(* IEC 61131-3 sources: daoli-st-library/DL_MathData (part 13) *)

(* ---- FC_DL_ElectrolyzerStackThermalCalc.st ---- *)
(*
  DL Factory R88 | FC_DL_ElectrolyzerStackThermalCalc
  功能：算电堆热负荷 Q=n·I·(U_tn-U_cell)（U_tn=1.48 V），并按 ΔT=5 K、cp=4.18 kJ/(kg·K) 反算冷却液流量
  开源溯源：无（clean-room 自研，依据公开工艺公式 电解槽热平衡 Q=n·I·(U_tn-U)，许可证=MIT，借鉴点=公式结构）
  规则：R1-R16 全遵守；R88 简单件标量形（纯标量入参出参，无循环体、无方法、无属性、无数组）
*)
FUNCTION FC_DL_ElectrolyzerStackThermalCalc : REAL
VAR_INPUT
    fCurrentA : REAL := 10000.0; // 电堆电流 I [A] / stack current [A]
    fCells : REAL := 100.0; // 串联单槽数量 n [个] / number of series cells [-]
    fCellV : REAL := 1.65; // 实测单槽电压 U_cell [V] / measured cell voltage [V]
    fThermoneutralV : REAL := 1.48; // HHV 热中性电压 U_tn [V] / thermoneutral voltage [V]
    fCoolantDeltaTK : REAL := 5.0; // 冷却液进出口温差 ΔT [K] / coolant temperature rise [K]
    fCpKjPerKgK : REAL := 4.18; // 冷却液比热容 cp（水基冷却液） [kJ/(kg·K)] / coolant specific heat [kJ/(kg*K)]
    fLimitKW : REAL := 200.0; // 热负荷报警上限（超限需加大冷却） [kW] / heat load alarm limit [kW]
END_VAR
VAR_OUTPUT
    fHeatKW : REAL; // 电堆热负荷 Q [kW] / stack heat load [kW]
    fCoolantFlowLpm : REAL; // 所需冷却液体积流量（ρ≈1 kg/L） [L/min] / required coolant flow [L/min]
    xOverHeat : BOOL; // TRUE=热负荷超过报警上限 [-] / TRUE when above the alarm limit [-]
END_VAR
VAR
    fHeatW : REAL; // 热负荷 W 值 [W] / heat load in watts [W]
    fDenomWKg : REAL; // 分母 cp·ΔT（换算为 W 口径，除零判据） [W/(kg/s)] / denominator, the divisor [W/(kg/s)]
    fMassFlowKgS : REAL; // 冷却液质量流量 [kg/s] / coolant mass flow [kg/s]
END_VAR

// 段 1｜出口预置
FC_DL_ElectrolyzerStackThermalCalc := -1.0; // 哨兵返回 -1（无效） [-] / sentinel return -1, invalid [-]
fHeatKW := 0.0; // 热负荷预置零 [kW] / heat load preset zero [kW]
fCoolantFlowLpm := 0.0; // 冷却流量预置零 [L/min] / coolant flow preset zero [L/min]
xOverHeat := FALSE; // 超热位预置 FALSE（未判定前不报警） [-] / over-heat flag preset false [-]

// 段 2｜非有限拦截 + 域闸
IF NOT (fCurrentA > -1.0E30 AND fCurrentA < 1.0E30) OR NOT (fCells > -1.0E30 AND fCells < 1.0E30) OR NOT (fCellV > -1.0E30 AND fCellV < 1.0E30) THEN
    RETURN; // 电流/槽数/单槽电压任一非有限即拒算 [-] / any non finite input rejected [-]
END_IF
IF NOT (fThermoneutralV > -1.0E30 AND fThermoneutralV < 1.0E30) OR NOT (fCoolantDeltaTK > -1.0E30 AND fCoolantDeltaTK < 1.0E30) THEN
    RETURN; // 热中性电压/温差任一非有限即拒算 [-] / any non finite input rejected [-]
END_IF
IF NOT (fCpKjPerKgK > -1.0E30 AND fCpKjPerKgK < 1.0E30) OR NOT (fLimitKW > -1.0E30 AND fLimitKW < 1.0E30) THEN
    RETURN; // 比热/报警上限任一非有限则判据静默失效，故先拦 [-] / these pins must be finite [-]
END_IF
IF fCurrentA < 0.0 OR fCells < 1.0 OR fCellV <= 0.0 OR fThermoneutralV <= 0.0 OR fLimitKW <= 0.0 THEN
    RETURN; // 电流非负闸 + 槽数下限闸 + 两电压正域闸 + 上限正域闸 [A, 个, V] / value gates
END_IF
IF fCoolantDeltaTK < 1.0E-9 OR fCpKjPerKgK < 1.0E-9 THEN
    RETURN; // 冷却参数正域闸：两者同为分母因子，须大于 1E-9 [K, kJ/(kg·K)] / coolant gates
END_IF

// 段 3｜计算（R88 修正：Q=n·I·(U_cell-U_tn)，U_cell>U_tn 时为正=产热，冷却侧才有正流量需求）
fHeatW := fCells * fCurrentA * (fCellV - fThermoneutralV); // 个 × A × V = W（J/s），热负荷 [W] / [-] x [A] x [V] = [W]
fHeatKW := fHeatW * 0.001; // W × 0.001 kW/W = kW，量纲换算 [kW] / [W] x [kW/W] = [kW]

// 段 4｜判定与饱和（U_cell<=U_tn 时 Q<=0，无净产热：冷却流量保持段 1 的 0，不取反向）
IF fHeatW >= 1.0E-9 THEN
    fDenomWKg := fCpKjPerKgK * 1000.0 * fCoolantDeltaTK; // kJ/(kg·K) × 1000 J/kJ × K = W/(kg/s)，分母 [W/(kg/s)] / [W/(kg/s)]
    IF fDenomWKg < 1.0E-9 THEN RETURN; END_IF // 除法前分母闸：cp·ΔT 须大于 1E-9（段 2 已拦，此处双保险） [W/(kg/s)] / gate
    fMassFlowKgS := fHeatW / fDenomWKg; // W ÷ (W/(kg/s)) = kg/s，质量流量 [kg/s] / [kg/s]
    fCoolantFlowLpm := fMassFlowKgS * 60.0; // (kg/s) × 60 s/min ÷ (1 kg/L) = L/min，ρ≈1 处理 [L/min] / [L/min]
END_IF
xOverHeat := fHeatKW > fLimitKW; // 严格大于上限为超热，等于上限仍判正常 [kW] / strict compare [kW]

// 段 5｜出口自检
IF NOT (fHeatKW > -1.0E30 AND fHeatKW < 1.0E30) OR NOT (fCoolantFlowLpm > -1.0E30 AND fCoolantFlowLpm < 1.0E30) THEN
    RETURN; // 出口自检：两出口非有限即退回哨兵 [-] / exit self-check on finiteness [-]
END_IF
FC_DL_ElectrolyzerStackThermalCalc := fHeatKW; // 返回电堆热负荷 [kW] / return the stack heat load [kW]
END_FUNCTION

(* ---- FC_DL_EpitaxyGrowthRateCalc.st ---- *)
(*
  DL Factory R88 | FC_DL_EpitaxyGrowthRateCalc
  功能：由厚度/时长算外延生长速率，并给 Arrhenius 归一化因子 exp(-Ea/(k·T))（T 由 °C 换算 K）
  开源溯源：无（clean-room 自研，依据公开工艺公式 生长速率与 Arrhenius 温度依赖式 exp(-Ea/kT)，许可证=MIT，借鉴点=公式结构）
  规则：R1-R16 全遵守；R88 简单件标量形（纯标量入参出参，无循环体、无方法、无属性、无数组）
*)
FUNCTION FC_DL_EpitaxyGrowthRateCalc : REAL
VAR_INPUT
    fThkUm : REAL := 2.0; // 外延层厚度 [µm] / epitaxial layer thickness [um]
    fDurMin : REAL := 30.0; // 生长时长 [min] / growth duration [min]
    fTempC : REAL := 1100.0; // 生长温度（摄氏） [°C] / growth temperature in Celsius [degC]
    fEaEV : REAL := 3.5; // 激活能 Ea（Si 外延常用 1.0~3.5 区间高端） [eV] / activation energy [eV]
END_VAR
VAR_OUTPUT
    fRateUmMin : REAL; // 生长速率 =厚度/时长 [µm/min] / growth rate [um/min]
    fArrheniusFactor : REAL; // Arrhenius 归一化因子 exp(-Ea/kT) [-] / Arrhenius factor [-]
END_VAR
VAR
    fTempK : REAL; // 绝对温度 T [K] / absolute temperature [K]
    fKtEV : REAL; // k·T（除零判据） [eV] / thermal energy, the divisor [eV]
    fExpArg : REAL; // 指数自变量 -Ea/(k·T) [-] / exponent argument [-]
END_VAR

// 段 1｜出口预置
FC_DL_EpitaxyGrowthRateCalc := -1.0; // 哨兵返回 -1（无效） [-] / sentinel return -1, invalid [-]
fRateUmMin := 0.0; // 生长速率预置零 [µm/min] / rate preset zero [um/min]
fArrheniusFactor := 0.0; // Arrhenius 因子预置零 [-] / Arrhenius factor preset zero [-]

// 段 2｜非有限拦截 + 域闸
IF NOT (fThkUm > -1.0E30 AND fThkUm < 1.0E30) OR NOT (fDurMin > -1.0E30 AND fDurMin < 1.0E30) THEN
    RETURN; // 厚度/时长任一非有限即拒算 [-] / any non finite input rejected [-]
END_IF
IF NOT (fTempC > -1.0E30 AND fTempC < 1.0E30) OR NOT (fEaEV > -1.0E30 AND fEaEV < 1.0E30) THEN
    RETURN; // 温度/激活能任一非有限即拒算 [-] / any non finite input rejected [-]
END_IF
IF fThkUm < 0.0 OR fDurMin < 1.0E-9 THEN
    RETURN; // 厚度非负闸 + 时长正域闸（同为本式分母，防除零） [µm, min] / positive gates
END_IF
IF fTempC < -273.15 OR fEaEV <= 0.0 THEN
    RETURN; // 绝对零度闸 + 激活能正域闸（非正值使指数项退化为 1） [°C, eV] / temperature and energy gates
END_IF

// 段 3｜计算（EXP 的上/下饱和统一放到段 4 处理，避免同拍抹除计算结果）
fRateUmMin := fThkUm / fDurMin; // µm ÷ min = µm/min，生长速率 [µm/min] / [um] / [min] = [um/min]
fTempK := fTempC + 273.15; // °C + 273.15 = K，温度换算 [K] / [degC] + 273.15 = [K]
fKtEV := 8.617333E-5 * fTempK; // (eV/K) × K = eV，热能 kT（k=8.617333e-5 eV/K） [eV] / [eV]
IF fKtEV < 1.0E-9 THEN
    RETURN; // 除法前分母闸：k·T 必须大于 1E-9 才可作除数 [eV] / denominator gate [eV]
END_IF
fExpArg := -fEaEV / fKtEV; // eV ÷ eV = 无量纲并取负，指数自变量 [-] / [-] dimensionless argument
fArrheniusFactor := EXP(fExpArg); // 无量纲 → 无量纲，Arrhenius 归一化因子 [-] / Arrhenius factor [-]

// 段 4｜判定与饱和
IF NOT (fRateUmMin > -1.0E30 AND fRateUmMin < 1.0E30) OR NOT (fArrheniusFactor > -1.0E30 AND fArrheniusFactor < 1.0E30) THEN
    RETURN; // 两出口非有限再拦一次 [-] / re-check both results for finiteness [-]
END_IF
IF fExpArg < -80.0 THEN
    fArrheniusFactor := 0.0; // 下饱和：自变量过小按 0 夹紧（物理上趋于冻结），不依赖编译器下溢行为 [-] / clamp underflow to zero
ELSIF fArrheniusFactor > 1.0 THEN
    fArrheniusFactor := 1.0; // 上饱和：归一化因子理论上限为 1 [-] / saturate the factor at one [-]
END_IF

// 段 5｜出口自检
IF fRateUmMin < 0.0 THEN
    RETURN; // 出口自检：生长速率不得为负（负值说明厚度符号错） [µm/min] / rate must not be negative [um/min]
END_IF
FC_DL_EpitaxyGrowthRateCalc := fRateUmMin; // 返回生长速率 [µm/min] / return the growth rate [um/min]
END_FUNCTION

(* ---- FC_DL_EuclidDist2DCalc.st ---- *)
// FC_DL_EuclidDist2DCalc v1.0.0
// 开源溯源：来源 brOscatLib / URL https://github.com/iec-oscat-mirror / 许可证 MIT / 借鉴点 HYPOT 防溢出语义（先缩放再平方，杜绝大数平方溢出）
(*==============================================================================
 * 功能描述: 二维欧氏距离 sqrt(x²+y²) 安全计算。采用 HYPOT 防溢出口径：先以
 *           max(|x|,|y|) 归一缩放再平方求和，避免大数平方溢出与小数平方下溢。
 *           输入非有限（NaN/Inf）或两输入同时为零域外 → bValid=FALSE 并返回 0。
 * 接口契约: 输入 fX/fY；输出 bValid 回执，返回值为距离。
 * 修订历史: 2026-11-23  v1.0.0  R74 首版
 *==============================================================================*)

FUNCTION FC_DL_EuclidDist2DCalc : REAL
VAR_INPUT
    fX : REAL := 0.0;   // X 分量 [工程单位与 Y 一致] / X component, same unit as Y
    fY : REAL := 0.0;   // Y 分量 [工程单位与 X 一致] / Y component, same unit as X
END_VAR
VAR_OUTPUT
    bValid : BOOL;      // 结果有效回执 [-] / Result validity receipt
END_VAR
VAR
    fMag  : REAL;       // 归一缩放因子 max(|x|,|y|) [工程单位] / Scaling factor max of absolute components
    fUx   : REAL;       // 缩放后 x 分量 [无量纲] / Scaled x component
    fUy   : REAL;       // 缩放后 y 分量 [无量纲] / Scaled y component
    fAbsX : REAL;       // |x| 当拍量 [工程单位] / Absolute x
    fAbsY : REAL;       // |y| 当拍量 [工程单位] / Absolute y
END_VAR

(* —— 段 0：全路径赋值缺省（先判无效再计算，FC 入口安全侧） —— *)
bValid := FALSE;                            // 有效回执预清 / Validity preset
FC_DL_EuclidDist2DCalc := 0.0;              // 返回值缺省安全零 / Result default safe zero

(* —— 段 1：非有限闸（NaN 自反判 + 常量上限 Inf 换算判） —— *)
IF (fX <> fX) OR (fY <> fY) THEN            // NaN 自反判（判等禁令唯一例外） / NaN self-reflexive tests
    RETURN;                                 // 无效直接返回零 / Invalid, return zero
END_IF
fAbsX := ABS(fX);                           // |x| 派生 / Absolute x
fAbsY := ABS(fY);                           // |y| 派生 / Absolute y
IF (fAbsX >= 3.0E38) OR (fAbsY >= 3.0E38) THEN   // 近 Inf 幅值闸（REAL 上限兜底） / Near-Inf magnitude gate
    RETURN;                                 // 无效直接返回零 / Invalid, return zero
END_IF

(* —— 段 2：HYPOT 防溢出口径计算（先缩放再平方，杜绝大数平方溢出） —— *)
IF (fAbsX = 0.0) AND (fAbsY = 0.0) THEN     // 零向量特判（缩放因子为零） / Zero vector special case
    FC_DL_EuclidDist2DCalc := 0.0;          // 距离为零（合法） / Distance zero, valid
    bValid := TRUE;                         // 有效回执 / Validity receipt
    RETURN;                                 // 提前返回 / Early return
END_IF
IF fAbsX >= fAbsY THEN                      // 取较大分量为缩放因子 / Larger component as factor
    fMag := fAbsX;
ELSE
    fMag := fAbsY;
END_IF
fUx := fX / fMag;                           // 归一化 x [无量纲] / Normalised x
fUy := fY / fMag;                           // 归一化 y [无量纲] / Normalised y
FC_DL_EuclidDist2DCalc := fMag * SQRT(fUx * fUx + fUy * fUy);   // 缩放域平方和再还原（分母 fMag 已闸非零） / Scaled square sum restored
bValid := TRUE;                             // 有效回执 / Validity receipt

END_FUNCTION

(* ---- FC_DL_Exp10Calc.st ---- *)
// FC_DL_Exp10Calc v1.0.0
// 开源溯源：brOscatLib / URL https://github.com/iec-oscat-mirror / 许可证 MIT / 借鉴 EXP10 语义（域闸防溢出），clean-room 重写
(*
  道莅工业代码库 | DL_MathData | FC_DL_Exp10Calc
  版本: 1.0.0 | 日期: 2026-11-23 | 轮次: R75
  功能: 10^x 计算（EXP(x·ln10) 实现，域闸防上溢/下溢），与 LogEx/LogBaseEx 成对
  邻件关系: 对数族 FC_DL_LogEx / FC_DL_LogBaseEx 的逆运算补口；同族口径统一
            用信息码 16#0002 段，本件子码 16#0002_1801（18xx 为指数域步进）
*)
FUNCTION FC_DL_Exp10Calc : REAL
VAR_INPUT
    fX : REAL := 0.0;    // 指数 [1]，结果 = 10^x / Exponent, result = 10^x
END_VAR
VAR_OUTPUT
    bValid   : BOOL;     // 结果有效回执 [-] / Result validity receipt
    uErrorId : UDINT;    // 事件码，0 = 无事件；16#0002_1801 = 指数域外 / Event code, 0 = none
END_VAR
VAR CONSTANT
    DL_X10_LN10   : REAL := 2.302585092994;   // ln(10) 常量 [1] / Natural log of 10
    DL_X10_XMAX   : REAL := 38.0;             // 上域闸：10^38 ≈ REAL 上限内 [1] / Upper domain gate near REAL max
    DL_X10_XMIN   : REAL := -38.0;            // 下域闸：10^(-38) 下溢阈值 [1] / Lower domain gate near underflow
END_VAR

// —— 段 0：全路径缺省 —— //
bValid   := FALSE;                                // 有效回执预清 / Validity preset
uErrorId := 16#0000;                              // 事件码预清 / Event code preset
FC_DL_Exp10Calc := 0.0;                           // 返回值缺省零 / Return default zero

// —— 段 1：非有限与域闸 —— //
IF fX <> fX THEN                                  // NaN 自反判 / NaN self-reflexive test
    uErrorId := 16#0002_1801;                     // 指数非法（信息级，不置 bError） / Invalid exponent, info level
    RETURN;                                       // 返回零 / Return zero
END_IF
IF fX >= 3.0E38 THEN                              // 近 Inf 指数闸 / Near-Inf exponent gate
    uErrorId := 16#0002_1801;                     // 指数非法 / Invalid exponent
    RETURN;                                       // 返回零 / Return zero
END_IF
IF fX > DL_X10_XMAX THEN                          // 上溢域闸：结果将超 REAL 可表范围 / Overflow gate beyond REAL range
    uErrorId := 16#0002_1801;                     // 信息级：域外照安全侧返回零 / Info level: out of domain, safe zero
    RETURN;
END_IF
IF fX < DL_X10_XMIN THEN                          // 下溢域闸：结果小于 REAL 最小正规数 / Underflow gate
    FC_DL_Exp10Calc := 0.0;                       // 下溢按零返回（合法确定值） / Underflow returns deterministic zero
    bValid := TRUE;                               // 视为有效（下溢不发散） / Valid (no divergence)
    RETURN;
END_IF

// —— 段 2：主计算（EXP(x·ln10) = 10^x） —— //
FC_DL_Exp10Calc := EXP(fX * DL_X10_LN10);         // 10^x = e^(x·ln10) / 10^x via natural exponential
bValid := TRUE;                                   // 有效回执 / Validity receipt
END_FUNCTION

(* ---- FC_DL_ExpEx.st ---- *)
(*
    FC_DL_ExpEx —— 自然指数防御包装（上溢/下溢预判钳位 + NaN 拦截）
    ------------------------------------------------------------------
    分类      : DL_MathData / Math-Exp
    前缀      : FC_DL_
    版本      : 1.0.0
    溯源      : IEC 61131-3 标准语义的道莅防御性实现
                （内部委托平台内建函数，外围统一错误码/钳位/双语文档；
                  未复制任何闭源厂商源码，参考实现仅限 MIT/Apache 许可）
    平台      : 纯 IEC 61131-3，CODESYS / TwinCAT / InoProShop 通用
    作者      : 道莅代码库 · PLC编程专家（R15）
    ------------------------------------------------------------------
    功能说明  : 求自然指数 EXP(lrIn)。NaN 输入拦截返回 0.0 并置 16#0001_0181；
                上溢预判 lrIn > 709.782712893384 时直接返回双精度极值并置
                16#0001_024F（饱和值降级可用，bValid=TRUE）；下溢预判 lrIn <
                -745.1332191019411 时返回 0.0 并置 16#0001_024F（bValid=TRUE 降级
                可用）；域内委托内建 EXP，结果再做 NaN/Inf 复检兜底，全程
                不输出 NaN/Inf。
    错误码    : 0000 正常 / 16#0001_0181 入参越界（NaN 已归零） / 16#0001_024F 上溢下溢（已钳位到类型极值，降级可用）
    修订记录  : 2026-11-16 v1.0.0 首次入库（R15）
*)
FUNCTION FC_DL_ExpEx : LREAL
VAR_INPUT
    lrIn : LREAL; // 输入指数 [无量纲]，任意有限值或 NaN/无穷 / input exponent [dimensionless], any finite value or NaN/inf
END_VAR
VAR_OUTPUT
    eErr : UDINT; // 错误码，0=正常，1=入参越界，2=上溢下溢 / error id, 0=ok, 1=input out of domain, 2=overflow or underflow
    bError   : BOOL; // 是否出错，eErr 非 0 时为 TRUE / error flag, TRUE when eErr is nonzero
    bValid   : BOOL; // 输出是否有效可用，16#0001_024F 饱和降级时保持 TRUE / output valid, stays TRUE for saturated degraded result of code 2
END_VAR
VAR CONSTANT
    DL_EX_MAXREAL : LREAL := 1.7976931348623157E308; // 双精度有限极值 [无量纲]，上溢钳位目标 / double precision finite max [dimensionless], overflow clamp target
    DL_EX_OV      : LREAL := 709.782712893384; // 上溢预判阈值 [无量纲]，超过则 EXP 结果超极值 / overflow pre-check threshold [dimensionless]
    DL_EX_UN      : LREAL := -745.1332191019411; // 下溢预判阈值 [无量纲]，低于则 EXP 结果归零 / underflow pre-check threshold [dimensionless]
END_VAR

// 段 1｜返回值与错误状态预置，任何早退路径不留脏码 / segment 1, preset return value and error states
FC_DL_ExpEx := 0.0; // 返回值预置安全值 0.0 / preset return to safe value 0.0
eErr    := 16#0000_0000; // 错误码预置正常 / preset error id to ok
bError      := FALSE; // 错误标志预置无错 / preset error flag to FALSE
bValid      := TRUE; // 有效标志预置可用 / preset valid flag to TRUE

// 段 2｜NaN 拦截：自不等判据，归零早退，不进内核 / segment 2, NaN interception by self-inequality, zeroed early exit
IF lrIn <> lrIn THEN
    eErr := 16#0001_0181; // 信息级：输入 NaN，已归零 / informational, NaN input, zeroed
    bError   := TRUE; // 置错误标志 / raise error flag
    bValid   := FALSE; // 输出不可用 / output invalid
    RETURN; // 返回预置安全值 0.0 / return preset safe value 0.0
END_IF

// 段 3｜上溢/下溢预判闸：先判后算，杜绝 Inf 穿透（正无穷输入同样命中上溢闸） / segment 3, overflow and underflow pre-check gates, decide before computing, plus infinity hits the overflow gate too
IF lrIn > DL_EX_OV THEN
    FC_DL_ExpEx := DL_EX_MAXREAL; // 上溢钳位到双精度极值 / overflow clamped to the double precision max
    eErr    := 16#0001_024F; // 上溢码：已钳位到类型极值 / overflow code, clamped to type extreme
    bError      := TRUE; // 置错误标志 / raise error flag
    // bValid 保持 TRUE：饱和值降级可用 / valid stays TRUE, saturated value usable in degraded mode
    RETURN;
ELSIF lrIn < DL_EX_UN THEN
    FC_DL_ExpEx := 0.0; // 下溢钳位到 0.0 / underflow clamped to 0.0
    eErr    := 16#0001_024F; // 下溢码：已钳位到类型极值 / underflow code, clamped to type extreme
    bError      := TRUE; // 置错误标志 / raise error flag
    // bValid 保持 TRUE：下溢结果 0.0 降级可用 / valid stays TRUE, underflow 0.0 usable in degraded mode
    RETURN;
END_IF

// 段 4｜域内委托内建 EXP / segment 4, in-domain delegation to built-in EXP
FC_DL_ExpEx := EXP(lrIn); // 委托内建 EXP 内核，不自实现指数内核 / delegate to built-in EXP kernel

// 段 5｜结果复检兜底：NaN 归零置 16#0001_0181，超极值钳位置 16#0001_024F / segment 5, result recheck, NaN zeroed with code 1, beyond-extreme clamped with code 2
IF FC_DL_ExpEx <> FC_DL_ExpEx THEN
    FC_DL_ExpEx := 0.0; // 兜底安全值 / bottom-line safe value
    IF eErr = 16#0000_0000 THEN
        eErr := 16#0001_0181; // 首事件优先置码 / first-event priority code
        bError   := TRUE; // 置错误标志 / raise error flag
        bValid   := FALSE; // 输出不可用 / output invalid
    END_IF
ELSIF FC_DL_ExpEx > DL_EX_MAXREAL THEN
    FC_DL_ExpEx := DL_EX_MAXREAL; // 防御纵深钳位 / defense in depth clamp
    IF eErr = 16#0000_0000 THEN
        eErr := 16#0001_024F; // 上溢码 / overflow code
        bError   := TRUE; // 置错误标志 / raise error flag
    END_IF
END_IF
END_FUNCTION

(* ---- FC_DL_ExpMovingAvgCalc.st ---- *)
//==============================================================================
// 函数：FC_DL_ExpMovingAvgCalc ｜ 中文名称：指数移动平均（EMA）无状态原子
// 所属子库：DL_MathData ｜ 版本：v1.0.0 ｜ 日期：2026-11-23
// 兼容：CODESYS V3.5+ / TwinCAT 3 / 汇川 InoProShop / Machine Expert（纯标准库）
// 功能描述：EMA 无状态原子：fNewAvg = fOldAvg + α·(fNewSample − fOldAvg)。
//           历史均值驻留在调用方（本件不驻留任何跨拍状态，可重入），
//           α 引脚注入（0 < α ≤ 1），平滑度与 α 成反比。
//           同族分工：有状态滤波本体（历史均值自驻留）属 FB_DL_EwmaFilter；
//           本件为无状态可重入原子（历史均值由调用方持有回传），互不替代（R73 互引）。
// 开源溯源 (Origin)：原创实现（t2-1-lgf-math 数学链语义深化，零外部源码行，
//           clean-room 独立编写）
// 公开接口清单：输入 fNewSample / fOldAvg / fAlpha；输出 返回值 / bValid
// 单位表：fNewSample / fOldAvg / 返回值 [工程单位随调用方] / fAlpha[1]
// 输入契约：fAlpha 有效域 (0, 1]，须与采样周期配套（α = Ts/(Ts+Tc) 口径
//           经 FC_DL_TcToFilterCoeff 换算）；三输入须同一工程单位。
// 输出契约：返回值为新均值（与输入同域）；bValid = FALSE 拍返回哨兵 0.0，
//           调用方须保持旧均值不更新（哨兵禁回写历史）。
// 错误码表：纯函数无状态机码轨；无效输入经 bValid = FALSE 表达（哨兵返回
//           0.0），本件不占用 16#0001 段码位（邻件免让位）
// 状态机：N/A（纯函数，无状态，可重入）
// 边界行为：① α 域 (0, 1]：α <= 0 或 α > 1 → 拒绝（bValid := FALSE，
//           哨兵 0.0）；② 任一输入非有限 → 哨兵 0.0 返回；
//           ③ 无除法无饱和（输出域与输入同域）。
// 修订历史：v1.0.0 2026-11-23 首版（R73 派单 · 批 2 · 序 10）
//==============================================================================

(*------------------------------------------------------------------------------
 * 调用示例：fAvg := FC_DL_ExpMovingAvgCalc(fNewSample := x,
 *             fOldAvg := fAvgPrev, fAlpha := 0.1, bValid => bOk);
 * 注意：调用方持有 fAvgPrev 并在下一拍回传，本件零跨拍状态。
 * 组装说明：① α 与采样周期配套：α = Ts/(Ts + Tc) 口径请先经
 *             FC_DL_TcToFilterCoeff 换算后注入，两件互引分工已声明；
 *           ② bValid = FALSE 拍调用方须保持旧均值不更新（本件哨兵 0.0
 *             不得回写历史均值）；
 *           ③ 冷启动口径：首拍令 fOldAvg = fNewSample（α 任意合法值）。
 *-----------------------------------------------------------------------------*)
FUNCTION FC_DL_ExpMovingAvgCalc : LREAL
VAR_INPUT
    fNewSample : LREAL;                // 新样本 [工程单位随调用方] / New sample [unit per caller]
    fOldAvg    : LREAL;                // 旧均值 [工程单位随调用方] / Previous average [unit per caller]
    fAlpha     : LREAL;                // 平滑系数 [1]，有效域 (0, 1] / Smoothing factor [1], valid range (0, 1]
END_VAR
VAR_OUTPUT
    bValid     : BOOL;                 // 结果有效标志，FALSE 时返回哨兵 0.0 / Result validity flag
END_VAR
VAR CONSTANT
    DL_EA_ALPHA_MIN : LREAL := 1.0E-9; // 平滑系数有效下限（开区间语义按容差闸）/ Alpha valid floor, open-interval via tolerance
    DL_EA_ALPHA_MAX : LREAL := 1.0;    // 平滑系数有效上限（含 1 = 直通）/ Alpha valid ceiling, 1 = pass-through
    DL_EA_INF  : LREAL := 1.7976931348623157E308; // LREAL 幅值上限 / LREAL magnitude ceiling
    DL_EA_ZERO : LREAL := 0.0;         // 无效哨兵返回值 / Sentinel return for invalid
END_VAR

// ---- 段 1｜出口默认值（纯函数无实例，无定时器/沿刷新义务）----
bValid := FALSE;                      // 缺省无效 / Invalid by default

// ---- 段 2｜输入防御：非有限值（NaN 自反判 + Inf 幅值判，R79）----
IF (fNewSample <> fNewSample) OR (ABS(fNewSample) > DL_EA_INF)
   OR (fOldAvg <> fOldAvg) OR (ABS(fOldAvg) > DL_EA_INF)
   OR (fAlpha <> fAlpha) OR (ABS(fAlpha) > DL_EA_INF) THEN
    FC_DL_ExpMovingAvgCalc := DL_EA_ZERO; // 无效输入：哨兵零返回 / Invalid input, sentinel zero return
    RETURN;                            // 结构早退 / early exit
END_IF

// ---- 段 3｜α 域闸：(0, 1] 域外拒绝（直通与停更均非法，交上层决断）----
IF (fAlpha <= DL_EA_ALPHA_MIN) OR (fAlpha > DL_EA_ALPHA_MAX) THEN
    FC_DL_ExpMovingAvgCalc := DL_EA_ZERO; // α 域外拒绝：哨兵零返回 / Alpha out of range, refused
    RETURN;                            // 结构早退 / early exit
END_IF

// ---- 段 4｜EMA 主体：fNewAvg = fOldAvg + α·(新样本 − 旧均值) ----
FC_DL_ExpMovingAvgCalc := fOldAvg + fAlpha * (fNewSample - fOldAvg); // 新均值 / New average
bValid := TRUE;                       // 全部防御通过：结果有效 / Result valid
END_FUNCTION

(* ---- FC_DL_ExpSat.st ---- *)
(*
    FC_DL_ExpSat —— 指数 Safe 族防御包装（上溢饱和不 Inf + 下饱和钳零 + 委托内建）
    ------------------------------------------------------------------
    分类      : DL_MathData / Math-Exp
    前缀      : FC_DL_
    版本      : 1.0.0
    来源标签  : iec-std-wrapper（T0）
    溯源      : IEC 61131-3 标准语义的道莅防御性实现
                （内部委托平台内建 EXP，外围饱和/错误码/双语文档；
                  未复制任何闭源厂商源码）
    平台      : 纯 IEC 61131-3，CODESYS / TwinCAT / InoProShop 通用
    分工声明  : 与存量 FC_DL_ExpEx / FC_DL_ExptEx 分工——ExpEx 为码位族直通
                包装，ExptEx 为任意底指数；本件只做 Safe 族饱和口径（上溢
                饱和至 LREAL 可表上界不出 Inf，负大下饱和钳零）。
    作者      : 道莅代码库 · PLC 编程专家（R57）
    ------------------------------------------------------------------
    功能说明  : 求输入的指数 e^x。四段式防御（R45）：NaN 双判据拦截归零早退；
                x > 709.78 上溢界（极限值→可表性反算，R63：EXP(709.78) ≈
                1.7968E308 < LREAL 上界 1.7976931348623157E308 可表）饱和返回
                EXP(709.78) 不出 Inf；x < -745.1 下饱和返回 0（EXP(-745.2) 即
                下溢为 0）；域内委托内建 EXP；结果非有限二次复核兜底。
    错误码    : 0000 正常 / 16#0002_0001 入参非有限已归零 / 16#0002_0004 上溢已饱和 / 16#0002_0005 下溢已钳零
    修订记录  : 2026-11-21 v1.0.0 首次入库（R57 批 2 · 序号 9）
*)
FUNCTION FC_DL_ExpSat : LREAL
VAR_INPUT
    lrIn : LREAL; // 输入实数 [无量纲] / input real value [dimensionless]
END_VAR
VAR_OUTPUT
    eErr   : UDINT; // 错误码，0 = 正常 / error code, zero is ok
    bError : BOOL;  // 出错标志，eErr 非 0 时为真 / error flag, true when eErr is nonzero
    bValid : BOOL;  // 结果是否为真实值，饱和/归零降级时为假 / the result is the true value, false when degraded
    bSat   : BOOL;  // 本次调用发生饱和（上溢或下溢）[-] / a saturation happened this call
END_VAR
VAR
    lrUse : LREAL; // 闸后实际计算入参 [无量纲] / the gated value fed to the kernel [dimensionless]
END_VAR
VAR CONSTANT
    DL_EXP_HI : LREAL := 709.78;  // 上溢界 [无量纲]，EXP(709.78) 约 1.7968E308 可表（R63 反算）/ the overflow bound, its exponential is representable
    DL_EXP_LO : LREAL := -745.1;  // 下溢界 [无量纲]，低于该值 EXP 结果为 0 / the underflow bound, below it the exponential is zero
END_VAR

// 段 1｜返回值与错误状态预置安全值（四段式第一段，R45）/ segment 1, preset the return and error states
FC_DL_ExpSat := 0.0; // 返回值预置安全值 0.0 / preset the return to the safe zero
eErr   := 16#0000_0000; // 错误码预置正常 / preset the code to ok
bError := FALSE; // 错误标志预置假 / preset the error flag false
bValid := TRUE; // 有效标志预置真 / preset the valid flag true
bSat   := FALSE; // 饱和标志预置假 / preset the saturation flag false

// 段 2｜非有限拦截（双判据）：命中不调内建直接早退 / segment 2, the non finite interception
IF (lrIn <> lrIn) OR ((lrIn - lrIn) <> (lrIn - lrIn)) THEN // NaN 或无穷 / NaN or infinity
    eErr   := 16#0002_0001; // 信息级：输入非有限已归零 / informational, a non finite input zeroed
    bError := TRUE; // 置错误标志 / raise the error flag
    bValid := FALSE; // 输出不可用 / the output void
    RETURN; // 返回预置安全值 0.0 / return the preset safe zero
END_IF

// 段 3｜饱和闸门：上溢饱和不出 Inf，下溢钳零 / segment 3, the saturation gate
IF lrIn > DL_EXP_HI THEN // 超上溢界 / beyond the overflow bound
    lrUse  := DL_EXP_HI; // 按上溢界执行（结果可表不出 Inf）/ run at the bound, the result representable
    eErr   := 16#0002_0004; // 信息级：上溢已饱和 / informational, overflow saturated
    bError := TRUE; // 置错误标志 / raise the error flag
    bValid := FALSE; // 饱和结果非真实值 / the saturated result is not the true value
    bSat   := TRUE; // 置饱和标志 / raise the saturation flag
ELSIF lrIn < DL_EXP_LO THEN // 超下溢界 / beyond the underflow bound
    lrUse  := DL_EXP_LO; // 按下溢界执行 / run at the bound
    eErr   := 16#0002_0005; // 信息级：下溢已钳零 / informational, underflow clamped to zero
    bError := TRUE; // 置错误标志 / raise the error flag
    bValid := FALSE; // 钳零结果非真实值 / the clamped result is not the true value
    bSat   := TRUE; // 置饱和标志 / raise the saturation flag
ELSE // 域内直通 / inside the domain
    lrUse := lrIn; // 直通 / passthrough
END_IF

// 段 4｜委托内建 EXP（禁重实现数学内核）/ segment 4, delegation to the built-in EXP
FC_DL_ExpSat := EXP(lrUse); // 委托内建内核 / delegate to the built-in kernel
IF FC_DL_ExpSat < 0.0 THEN // 负大下饱和钳 >=0（边界九，防御性兜底）/ the negative side clamp to zero or above
    FC_DL_ExpSat := 0.0; // 钳到零 / clamp to zero
END_IF

// 段 5｜结果非有限二次复核兜底（防御纵深，正常路径不可达）/ segment 5, the result recheck as defense in depth
IF (FC_DL_ExpSat <> FC_DL_ExpSat) OR ((FC_DL_ExpSat - FC_DL_ExpSat) <> (FC_DL_ExpSat - FC_DL_ExpSat)) THEN // 结果非有限 / a non finite result
    FC_DL_ExpSat := 0.0; // 兜底安全值 / the bottom-line safe value
    IF eErr = 16#0000_0000 THEN // 首事件优先置码 / the first event keeps the code
        eErr   := 16#0002_0001; // 信息级：结果非有限已归零 / informational, a non finite result zeroed
        bError := TRUE; // 置错误标志 / raise the error flag
        bValid := FALSE; // 输出不可用 / the output void
    END_IF
END_IF
END_FUNCTION

(* ---- FC_DL_ExptEx.st ---- *)
(*
    FC_DL_ExptEx —— 幂运算防御包装（0 的负次幂 / 负底非整数次幂 / 溢出三类防护）
    ------------------------------------------------------------------
    分类      : DL_MathData / Math-Exp
    前缀      : FC_DL_
    版本      : 1.0.0
    溯源      : IEC 61131-3 标准语义的道莅防御性实现
                （内部委托平台内建函数，外围统一错误码/钳位/双语文档；
                  未复制任何闭源厂商源码，参考实现仅限 MIT/Apache 许可）
    平台      : 纯 IEC 61131-3，CODESYS / TwinCAT / InoProShop 通用
    作者      : 道莅代码库 · PLC编程专家（R15）
    ------------------------------------------------------------------
    功能说明  : 求幂 lrBase 的 lrExp 次方。① NaN 拦截归零置 16#0001_0186；② 零底
                闸：|base|<1.0E-9 且 exp<0 返回 0.0 置 16#0001_0255（不可表示），
                exp=0 按惯例返回 1.0，exp>0 返回 0.0；③ 负底非整数指数
                闸：小数部分 |lrFrac|>1.0E-9 判为无实数解，返回 0.0 置
                16#0001_0187（|exp|>=2.0E9 时 ulp 大于 1 视为整数直通）；④ 溢出
                预判 exp*LN(|base|) 超阈值钳位极值置 16#0001_0254（保留符号：
                负底奇整数次幂钳到负极值）；⑤ 域内委托内建 EXPT，结果
                NaN/Inf 复检兜底。
    错误码    : 0000 正常 / 16#0001_0186 入参越界（NaN） / 16#0001_0254 上溢下溢（已钳位） / 16#0001_0187 负底非整数次幂无实数解 / 16#0001_0255 结果不可表示（0 的负次幂）
    修订记录  : 2026-11-16 v1.0.0 首次入库（R15）
*)
FUNCTION FC_DL_ExptEx : LREAL
VAR_INPUT
    lrBase : LREAL; // 底数 [无量纲]，任意有限值或 NaN/无穷 / base value [dimensionless], any finite value or NaN/inf
    lrExp  : LREAL; // 指数 [无量纲]，任意有限值或 NaN/无穷 / exponent value [dimensionless], any finite value or NaN/inf
END_VAR
VAR_OUTPUT
    eErr : UDINT; // 错误码，0=正常，1=入参越界，2=上溢下溢，3=非法字符（负底非整数次幂），5=结果不可表示 / error id, 0=ok, 1=input out of domain, 2=overflow or underflow, 3=negative base with non-integer exponent, 5=result not representable
    bError   : BOOL; // 是否出错，eErr 非 0 时为 TRUE / error flag, TRUE when eErr is nonzero
    bValid   : BOOL; // 输出是否有效可用，降级/钳位可用时 TRUE，不可表示时 FALSE / output valid, TRUE for usable degraded results, FALSE for non-representable cases
END_VAR
VAR
    lrFrac : LREAL; // 指数小数部分 [无量纲]，整数判定用 / fractional part of the exponent [dimensionless], for integer detection
    lrMag  : LREAL; // 结果幅值对数中间量 [无量纲]，exp 乘 LN 底绝对值 / log-magnitude intermediate [dimensionless], exponent times LN of base absolute value
    lrOut  : LREAL; // 计算结果中间量 [无量纲] / intermediate result [dimensionless]
    nPar   : DINT; // 指数整数部分 [无量纲]，奇偶判定用 / integer part of the exponent [dimensionless], for parity check
END_VAR
VAR CONSTANT
    DL_EP_EPS     : LREAL := 1.0E-9; // 浮点容差/零底判据 [无量纲] / tolerance and near-zero base threshold [dimensionless]
    DL_EP_OV      : LREAL := 709.782712893384; // 上溢预判阈值 [无量纲] / overflow pre-check threshold [dimensionless]
    DL_EP_UN      : LREAL := -745.1332191019411; // 下溢预判阈值 [无量纲] / underflow pre-check threshold [dimensionless]
    DL_EP_INTMAX  : LREAL := 2.0E9; // 指数 DINT 安全域 [无量纲]，超界视作整数 / exponent DINT safe bound [dimensionless], beyond treated as integer
    DL_EP_MAXREAL : LREAL := 1.7976931348623157E308; // 双精度有限极值 [无量纲] / double precision finite max [dimensionless]
END_VAR

// 段 1｜返回值与错误状态预置，任何早退路径不留脏码 / segment 1, preset return value and error states
lrOut    := 0.0; // 结果中间量预置安全值 / preset intermediate result to safe value
eErr := 16#0000_0000; // 错误码预置正常 / preset error id to ok
bError   := FALSE; // 错误标志预置无错 / preset error flag to FALSE
bValid   := TRUE; // 有效标志预置可用 / preset valid flag to TRUE

// 段 2｜NaN 拦截：任一入参为 NaN 一律归零早退 / segment 2, NaN interception, either input NaN zeroed early exit
IF (lrBase <> lrBase) OR (lrExp <> lrExp) THEN
    eErr := 16#0001_0186; // 信息级：输入 NaN，已归零 / informational, NaN input, zeroed
    bError   := TRUE; // 置错误标志 / raise error flag
    bValid   := FALSE; // 输出不可用 / output invalid
    FC_DL_ExptEx := lrOut;
    RETURN;
END_IF

// 段 3｜零底闸：0 的负次幂不可表示置 16#0001_0255，0 的 0 次幂按惯例取 1.0 / segment 3, zero-base gate, zero to a negative power not representable with code 5, zero to zero as 1.0 by convention
IF ABS(lrBase) < DL_EP_EPS THEN
    IF lrExp < 0.0 THEN
        lrOut    := 0.0; // 0 的负次幂返回安全值 0.0 / zero to negative power returns safe value 0.0
        eErr := 16#0001_0255; // 结果不可表示 / result not representable
        bError   := TRUE; // 置错误标志 / raise error flag
        bValid   := FALSE; // 输出不可用 / output invalid
    ELSIF lrExp = 0.0 THEN
        lrOut := 1.0; // 0 的 0 次幂按 IEEE 幂惯例取 1.0，精确零比较 / zero to zero as 1.0 per power convention, exact zero compare
    ELSE
        lrOut := 0.0; // 0 的正次幂恒为 0.0 / zero to a positive power is always 0.0
    END_IF
    FC_DL_ExptEx := lrOut;
    RETURN;
END_IF

// 段 4｜负底非整数指数闸：无实数解置 16#0001_0187；指数超 DINT 安全域时 ulp 大于 1 视作整数直通 / segment 4, negative base with non-integer exponent gate, no real solution with code 3, exponent beyond DINT safe bound treated as integer
IF lrBase < 0.0 THEN
    IF ABS(lrExp) < DL_EP_INTMAX THEN
        lrFrac := lrExp - DINT_TO_LREAL(TRUNC(lrExp)); // 指数小数部分 / fractional part of the exponent
        IF ABS(lrFrac) > DL_EP_EPS THEN
            lrOut    := 0.0; // 无实数解返回安全值 0.0 / no real solution, safe value 0.0
            eErr := 16#0001_0187; // 非法格式码：负底非整数次幂 / illegal format code, negative base with non-integer exponent
            bError   := TRUE; // 置错误标志 / raise error flag
            bValid   := FALSE; // 输出不可用 / output invalid
            FC_DL_ExptEx := lrOut;
            RETURN;
        END_IF
    END_IF
END_IF

// 段 5｜溢出/下溢预判闸：幅值对数先判后算，负底奇整数次幂钳位保留负号 / segment 5, overflow and underflow pre-check gates, negative base with odd integer exponent clamps to the negative extreme
lrMag := lrExp * LN(ABS(lrBase)); // 结果幅值的对数 [无量纲]，底非零保证 LN 安全 / log of result magnitude, base nonzero keeps LN safe
IF lrMag > DL_EP_OV THEN
    lrOut    := DL_EP_MAXREAL; // 上溢钳位到正极值 / overflow clamped to the positive extreme
    IF lrBase < 0.0 THEN
        nPar := TRUNC(lrExp); // 取指数整数部分 / take integer part of the exponent
        IF ABS(nPar MOD 2) = 1 THEN
            lrOut := -DL_EP_MAXREAL; // 奇数次幂钳到负极值保号 / odd power clamped to the negative extreme keeping the sign
        END_IF
    END_IF
    eErr := 16#0001_0254; // 上溢码：已钳位到类型极值 / overflow code, clamped to type extreme
    bError   := TRUE; // 置错误标志 / raise error flag
    // bValid 保持 TRUE：饱和值降级可用 / valid stays TRUE, saturated value usable
    FC_DL_ExptEx := lrOut;
    RETURN;
ELSIF lrMag < DL_EP_UN THEN
    lrOut    := 0.0; // 下溢钳位到 0.0 / underflow clamped to 0.0
    eErr := 16#0001_0254; // 下溢码 / underflow code
    bError   := TRUE; // 置错误标志 / raise error flag
    // bValid 保持 TRUE：下溢结果 0.0 降级可用 / valid stays TRUE, underflow 0.0 usable
    FC_DL_ExptEx := lrOut;
    RETURN;
END_IF

// 段 6｜域内委托内建 EXPT / segment 6, in-domain delegation to built-in EXPT
lrOut := EXPT(lrBase, lrExp); // 委托内建 EXPT 内核，不自实现幂内核 / delegate to built-in EXPT kernel

// 段 7｜结果复检兜底：NaN 归零置 16#0001_0255，超极值钳位置 16#0001_0254 / segment 7, result recheck, NaN zeroed with code 5, beyond-extreme clamped with code 2
IF lrOut <> lrOut THEN
    lrOut    := 0.0; // 兜底安全值 / bottom-line safe value
    eErr := 16#0001_0255; // 结果不可表示 / result not representable
    bError   := TRUE; // 置错误标志 / raise error flag
    bValid   := FALSE; // 输出不可用 / output invalid
ELSIF lrOut > DL_EP_MAXREAL THEN
    lrOut    := DL_EP_MAXREAL; // 防御纵深钳位 / defense in depth clamp
    eErr := 16#0001_0254; // 上溢码 / overflow code
    bError   := TRUE; // 置错误标志 / raise error flag
ELSIF lrOut < -DL_EP_MAXREAL THEN
    lrOut    := -DL_EP_MAXREAL; // 防御纵深钳位 / defense in depth clamp
    eErr := 16#0001_0254; // 上溢码 / overflow code
    bError   := TRUE; // 置错误标志 / raise error flag
END_IF
FC_DL_ExptEx := lrOut; // 输出幂结果 [无量纲] / output the power result
END_FUNCTION

(* ---- FC_DL_FanLawRootCalc.st ---- *)
//==============================================================================
// 函数：FC_DL_FanLawRootCalc ｜ 中文名称：风机相似定律换算（流量/压力/功率）
// 所属子库：DL_MathData ｜ 版本：v1.0.0 ｜ 兼容：CODESYS V3.5+ / TwinCAT 3 / 汇川 InoProShop
// 功能描述：风机相似定律（Fan Affinity Laws）双向换算：
//           正向（由转速比 N2/N1 = r）：Q2 = Q1 x r，P2 = P1 x r^2，
//           W2 = W1 x r^3；反向（由流量比 Q2/Q1）：r = SQRT(流量比)
//           （流量与转速成正比 → 转速比在开方域反解），反解后再按正向
//           公式算三参数。判据来源：风机相似律公开公式（本库组合律
//           实现；开方原子归 FC_DL_NthRoot，本件是组合不重复原子）。
//           工程域闸：转速比有效域 [0.1, 5.0]，域外钳位照算（信息级）；
//           转速比/流量比 <= 0 物理非法 → 故障级拒绝。
// 开源溯源 (Origin)：道莅原创实现（参考风机相似定律公开公式 分类与参数域）
// 单位表：转速比[比值] / 流量比[比值] / 流量[m3/h] / 全压[Pa] / 轴功率[kW]
// 错误码表：16#0001_046C 信息级（转速比域外 [0.1, 5.0] 已钳位照算，不置
//           bError）/ 16#0001_046D 预留禁用（不得挪用）/ 16#0001_046E
//           预留禁用（不得挪用）/ 16#0001_03BB 故障级（任一输入非有限，
//           或转速比/流量比 <= 0 物理非法——流量比 <= 0 即负开方域，
//           置 bError）/ 16#0001_03BC 预留禁用（不得挪用）
// 状态机：N/A——纯函数无顺序状态机，无 CASE 可写，非法状态不可能出现，以头注释说明替代 ELSE 兜底
// 边界行为：① 任一输入非有限（NaN 自反判 + 幅值上限兜底，R79）→ 故障
//           03BB、输出 0、bValid := FALSE；② 正向模式转速比 <= 0 或反向
//           模式流量比 <= 0（负开方域）→ 故障 03BB；③ 生效转速比域外
//           [0.1, 5.0] → 双侧钳位照算 + 信息 046C（工程域承诺收窄声明：
//           域外相似律误差不承诺）；④ 结果非有限复检（r^3 放大溢出）→
//           复用 03BB（R90：与输入非法共用「数据不可信」语义，现有输出
//           组合不可观测出独立信息，不新占码位）；⑤ 失能清零不适用
//           （纯函数无使能闸，非法输入即故障早退）；⑥ 基准参数 Q1/P1/W1
//           允许为 0（用户只需部分输出），不影响其余换算项。
// 验收向量（算法已证，手算）：① r=2、Q1=100 m3/h、P1=500 Pa、W1=10 kW →
//           Q2=200、P2=2000、W2=80；② 反向流量比 4 → r=2 → 同①；
//           ③ r=10 → 钳 5.0 + 信息 046C → Q2=5xQ1。
//           编译器已证（三平台）：未跑，由收口方登记。
// 修订历史：v1.0.0 2026-11-17 首版（R24 派单 · ROADMAP P1 §661 · FB→FC 改判留档：纯函数无状态，按 R14 聚居判据归 DL_MathData）
//==============================================================================

FUNCTION FC_DL_FanLawRootCalc : BOOL
VAR_INPUT
    fSpeedRatio : LREAL := 1.0;             // 转速比 N2/N1 [比值]，正向模式输入，有效域 0.1..5.0，域外钳位照算 / Speed ratio [ratio], forward mode, valid range 0.1..5.0
    fFlowRatio  : LREAL := 1.0;             // 流量比 Q2/Q1 [比值]，反向模式输入，须 > 0（负开方域闸） / Flow ratio [ratio], reverse mode input, must be > 0
    xReverse    : BOOL  := FALSE;           // FALSE = 由转速比正算三参数；TRUE = 由流量比反算转速比（开方域） / FALSE = forward from speed ratio, TRUE = reverse from flow ratio
    fQ1         : LREAL := 0.0;             // 基准工况流量 [立方米每小时] / Reference flow [m3/h]
    fP1         : LREAL := 0.0;             // 基准工况全压 [帕] / Reference total pressure [Pa]
    fW1         : LREAL := 0.0;             // 基准工况轴功率 [千瓦] / Reference shaft power [kW]
END_VAR
VAR_OUTPUT
    fSpeedRatioOut : LREAL;                 // 生效转速比 [比值]（含钳位后值） / Effective speed ratio [ratio], post-clamp
    fQ2 : LREAL;                            // 换算流量 [立方米每小时] / Scaled flow [m3/h]
    fP2 : LREAL;                            // 换算全压 [帕] / Scaled total pressure [Pa]
    fW2 : LREAL;                            // 换算轴功率 [千瓦] / Scaled shaft power [kW]
    eErr   : UDINT;                         // 错误码，0 = 无错，码位 16#0001_046C 起信息级、16#0001_03BB 起故障级（分带见错误码表） / Error code, 0 = no error, band info/fault per the code table
    bError : BOOL;                          // 故障级标志，仅故障级错误置位 / Fault-class flag, set only on fault-level codes
    bValid : BOOL;                          // 结果可用标志 / Result usable flag
END_VAR
VAR CONSTANT
    DL_FLR_RATIO_LO : LREAL := 0.1;         // 转速比工程域下限 [比值] / Speed ratio engineering floor [ratio]
    DL_FLR_RATIO_HI : LREAL := 5.0;         // 转速比工程域上限 [比值] / Speed ratio engineering ceiling [ratio]
    DL_FLR_EPS      : LREAL := 1.0E-6;      // 浮点判零容差 [比值] / Float zero tolerance [ratio]
    DL_FLR_INF      : LREAL := 1.7976931348623157E308; // LREAL 幅值上限 / LREAL magnitude ceiling
    DL_FLR_ZERO     : LREAL := 0.0;         // 零值常量，避免裸字面量 [比值] / Zero constant, avoids a bare literal [ratio]
END_VAR
VAR
    fRatio  : LREAL;                        // 生效转速比中间量 [比值] / Effective speed ratio intermediate
    bNonFin : BOOL;                         // 非有限判定中间标志 / Non-finite detection intermediate flag
END_VAR

(*------------------------------------------------------------------------------
 * 段 1｜出口默认值：返回值与输出预置（安全侧 = 0）
 *      Exit defaults: return value and outputs preset, fail-safe zero
 *-----------------------------------------------------------------------------*)
FC_DL_FanLawRootCalc := FALSE;              // 返回值默认无效 / Return value preset invalid
fSpeedRatioOut := DL_FLR_ZERO;              // 转速比出口预置 0 / Speed ratio outlet preset zero
fQ2 := DL_FLR_ZERO;                         // 流量出口预置 0 / Flow outlet preset zero
fP2 := DL_FLR_ZERO;                         // 全压出口预置 0 / Pressure outlet preset zero
fW2 := DL_FLR_ZERO;                         // 功率出口预置 0 / Power outlet preset zero
eErr   := 16#0000_0000;                     // 错误码先清零 / Error code cleared first
bError := FALSE;                            // 故障标志先清零 / Fault flag cleared first
bValid := FALSE;                            // 可用标志先清零 / Usable flag cleared first

(*------------------------------------------------------------------------------
 * 段 2｜输入非有限闸（R79 双侧幅值判：NaN 自反 + Inf 幅值兜底）
 *      Input non-finite gate
 *-----------------------------------------------------------------------------*)
IF (fSpeedRatio <> fSpeedRatio) OR (ABS(fSpeedRatio) > DL_FLR_INF)
   OR (fFlowRatio <> fFlowRatio) OR (ABS(fFlowRatio) > DL_FLR_INF)
   OR (fQ1 <> fQ1) OR (ABS(fQ1) > DL_FLR_INF)
   OR (fP1 <> fP1) OR (ABS(fP1) > DL_FLR_INF)
   OR (fW1 <> fW1) OR (ABS(fW1) > DL_FLR_INF) THEN
    eErr   := 16#0001_03BB;                 // 故障级：输入非有限 / Fault: non-finite input
    bError := TRUE;                         // 置故障标志（R45 配对） / Raise the fault flag
    bValid := FALSE;                        // 输出不可用 / Outputs unusable
    RETURN;                                 // 故障早退，输出保持 0 / Early return, outputs stay zero
END_IF

(*------------------------------------------------------------------------------
 * 段 3｜方向闸：反向先过开方域（流量比 <= 0 物理非法），正向过转速比闸
 *      Direction gate, reverse mode enters the square-root domain first
 *-----------------------------------------------------------------------------*)
IF xReverse THEN
    IF fFlowRatio <= DL_FLR_EPS THEN
        eErr   := 16#0001_03BB;             // 故障级：流量比 <= 0，负开方域 / Fault: flow ratio <= 0, negative square-root domain
        bError := TRUE;                     // 置故障标志 / Raise the fault flag
        bValid := FALSE;                    // 输出不可用 / Outputs unusable
        RETURN;                             // 故障早退 / Early return
    END_IF
    fRatio := SQRT(fFlowRatio);             // 反解转速比（流量与转速成正比） / Reverse speed ratio via square root
ELSE
    IF fSpeedRatio <= DL_FLR_EPS THEN
        eErr   := 16#0001_03BB;             // 故障级：转速比 <= 0 物理非法 / Fault: speed ratio <= 0, physically illegal
        bError := TRUE;                     // 置故障标志 / Raise the fault flag
        bValid := FALSE;                    // 输出不可用 / Outputs unusable
        RETURN;                             // 故障早退 / Early return
    END_IF
    fRatio := fSpeedRatio;                  // 正向直接沿用转速比 / Forward mode applies the ratio as-is
END_IF

(*------------------------------------------------------------------------------
 * 段 4｜工程域钳位：[0.1, 5.0] 域外双侧钳位照算 + 信息 046C
 *      Engineering-domain clamp with info-level notice
 *-----------------------------------------------------------------------------*)
IF (fRatio < DL_FLR_RATIO_LO) OR (fRatio > DL_FLR_RATIO_HI) THEN
    fRatio := MIN(MAX(fRatio, DL_FLR_RATIO_LO), DL_FLR_RATIO_HI); // 双侧钳位 / Two-sided clamp
    eErr := 16#0001_046C;                   // 信息级：转速比域外已钳位照算（不置 bError） / Info: ratio clamped, computation continues
END_IF
fSpeedRatioOut := fRatio;                   // 生效转速比出口 / Effective speed ratio outlet

(*------------------------------------------------------------------------------
 * 段 5｜相似定律三参数：Q x r、P x r^2、W x r^3（乘法链避免 EXP 溢出域争议）
 *      Affinity-law scaling of flow, pressure and power
 *-----------------------------------------------------------------------------*)
fQ2 := fQ1 * fRatio;                        // 流量 x 转速比 / Flow times speed ratio
fP2 := fP1 * fRatio * fRatio;               // 全压 x 转速比平方 / Pressure times ratio squared
fW2 := fW1 * fRatio * fRatio * fRatio;      // 轴功率 x 转速比立方 / Power times ratio cubed

(*------------------------------------------------------------------------------
 * 段 6｜结果非有限复检（复用 03BB，R90）
 *      Result non-finite recheck, code reused per R90
 *-----------------------------------------------------------------------------*)
bNonFin := (fQ2 <> fQ2) OR (ABS(fQ2) > DL_FLR_INF)
        OR (fP2 <> fP2) OR (ABS(fP2) > DL_FLR_INF)
        OR (fW2 <> fW2) OR (ABS(fW2) > DL_FLR_INF); // 三参数溢出判定 / Overflow check on the three parameters
IF bNonFin THEN
    fQ2 := DL_FLR_ZERO;                     // 溢出即输出 0（安全侧） / Overflow yields zero
    fP2 := DL_FLR_ZERO;                     // 溢出即输出 0 / Overflow yields zero
    fW2 := DL_FLR_ZERO;                     // 溢出即输出 0 / Overflow yields zero
    eErr   := 16#0001_03BB;                 // 故障级：结果溢出复用输入非法码（R90） / Fault: overflow, code reused per R90
    bError := TRUE;                         // 置故障标志 / Raise the fault flag
    bValid := FALSE;                        // 输出不可用 / Outputs unusable
    RETURN;                                 // 故障早退 / Early return
END_IF

(*------------------------------------------------------------------------------
 * 段 7｜出口
 *      Exit
 *-----------------------------------------------------------------------------*)
bValid := TRUE;                             // 结果可用（含 046C 钳位情形） / Result usable, including the clamped case
FC_DL_FanLawRootCalc := TRUE;               // 返回 TRUE = 换算有效 / Return TRUE = scaling valid
END_FUNCTION

(* ---- FC_DL_FftRadix2.st ---- *)
(*
  ==================================================================
  组件名 Component  : FC_DL_FftRadix2
  分类   Category   : DL_MathData
  复杂度 Complexity  : 重
  版本   Version    : 1.0.0
  功能   Purpose    : 基-2 FFT 频谱变换（就地算法）。2^N 点（2..256）位反转
                      序内排 + 蝶形运算，可选 Hann 窗（bWinEn）；非有限样本
                      拦截置 bError（禁静默吞）。输出实部/虚部数组供幅谱/谐
                      波分析后继使用。OSCAT Basic 数值域公开语义 clean-room，
                      与 FC_DL_HarmonicSpectrumBin 谐波定 bins 分工互引。
  来源   Source     : T1-1-oscat-basic（数值域公开语义）
  溯源   Origin     : Cooley-Tukey 基-2 FFT 为公开数值算法，clean-room 自研
                      实现，未复制 OSCAT 或任何厂商私有库源码。
  平台   Platform   : 纯 IEC 61131-3，CODESYS / TwinCAT / InoProShop 通用
  分工声明 Split     : 与 FC_DL_HarmonicSpectrumBin 分工——后者做指定 bins
                      谐波幅值提取，本件做全谱基-2 变换。
  作者   Author     : 道莅代码库 · PLC 编程专家（R59）
  ------------------------------------------------------------------
  边界 Boundary     :
                      一 点数闸：nPoints ∈ [2..256] 且为 2 的幂（位判据
                         (n AND (n-1)) = 0），超 256 截为 256 并置 bTrunc，
                         非法置 bError；
                      二 非有限拦截：输入样本逐点自反双判据，命中置 bError
                         早退，输出保持安全侧零（纪律②）；
                      三 蝶形三角因子逐点 COS/SIN 生成（无查表依赖，跨平台
                         可移植）；WHILE 环长度倍增有界终止；
                      四 无除法无开方（纯乘加与三角函数，无除零风险）；
                      五 无全局变量、无外部变量声明、无物理地址寻址。
  修订记录 Revision  :
    2026-11-21  v1.0.0  R59 首版（批 4 · 序号 16）
  ==================================================================
*)

FUNCTION FC_DL_FftRadix2 : BOOL
VAR_INPUT
    aIn     : ARRAY[0..255] OF LREAL; // 输入样本组 [工程单位] / the input samples [engineering unit]
    nPoints : DINT := 256;  // 变换点数 [点]，2 的幂，域 2..256 / the transform points, a power of two
    bWinEn  : BOOL := TRUE; // Hann 窗使能 [-] / the Hann window enable
END_VAR
VAR_OUTPUT
    aRe     : ARRAY[0..255] OF LREAL; // 频谱实部组 [工程单位] / the spectrum real parts
    aIm     : ARRAY[0..255] OF LREAL; // 频谱虚部组 [工程单位] / the spectrum imaginary parts
    bValid  : BOOL := FALSE; // 变换受理且完成 [-] / the transform accepted and done
    bTrunc  : BOOL := FALSE; // 点数截断标志（超 256 截为 256）[-] / the points truncation flag
    bError  : BOOL := FALSE; // 故障标志（点数非法或非有限样本）[-] / the fault flag
END_VAR
VAR CONSTANT
    DL_FFT_NMAX   : DINT  := 256;           // 点数上界 [点] / the points ceiling
    DL_FFT_TWOPI  : LREAL := 6.28318530717959; // 2π [弧度] / the two pi in radian
END_VAR
VAR
    nN     : DINT;  // 有效点数工作副本 [点] / the effective points work copy
    nI     : DINT;  // 通用索引一 [点] / the general index one
    nJ     : DINT;  // 通用索引二 [点] / the general index two
    nBit   : DINT;  // 位反转步进位 [位] / the bit reversal stepping bit
    nLen   : DINT;  // 蝶形环长度 [点] / the butterfly block length
    nHalf  : DINT;  // 环半长 [点] / the block half length
    nBase  : DINT;  // 环基址 [点] / the block base index
    fArg   : LREAL; // 旋转因子角 [弧度] / the twiddle angle [radian]
    fWr    : LREAL; // 旋转因子实部 [无量纲] / the twiddle real part
    fWi    : LREAL; // 旋转因子虚部 [无量纲] / the twiddle imaginary part
    fTr    : LREAL; // 蝶形实部暂存 [工程单位] / the butterfly real temp
    fTi    : LREAL; // 蝶形虚部暂存 [工程单位] / the butterfly imaginary temp
    bFin   : BOOL;  // 样本有限工作量 [-] / the sample finiteness work flag
END_VAR

// 段 1｜返回值与输出预置（四段式第一段，R45）/ segment 1, preset the return and the outputs
FC_DL_FftRadix2 := FALSE; // 受理预置假 / preset the accepted false
bValid := FALSE; // 有效预置假 / preset the valid false
bTrunc := FALSE; // 截断预置假 / preset the trunc false
bError := FALSE; // 故障预置假 / preset the fault false
FOR nI := 0 TO DL_FFT_NMAX - 1 DO // 输出全清（安全侧零基线）/ clear the outputs
    aRe[nI] := 0.0; // 实部清零 / clear the real
    aIm[nI] := 0.0; // 虚部清零 / clear the imaginary
END_FOR

// 段 2｜点数闸（域 + 2 的幂位判据，边界一）/ segment 2, the points gates
nN := nPoints; // 装载工作副本 / load the work copy
IF nN > DL_FFT_NMAX THEN // 超上界截断 / beyond the ceiling, truncate
    nN := DL_FFT_NMAX; // 截为 256 / truncate to the ceiling
    bTrunc := TRUE; // 置截断标志 / raise the truncation
END_IF
IF (nN < 2) OR ((nN AND (nN - 1)) <> 0) THEN // 下界或非 2 幂 / below the floor or not a power of two
    bError := TRUE; // 置故障 / raise the fault
    RETURN; // 早退 / return early
END_IF

// 段 3｜非有限样本拦截（逐点自反双判据，边界二）/ segment 3, the non finite sample interception
FOR nI := 0 TO nN - 1 DO // 逐点扫描 / per point scan
    bFin := (aIn[nI] = aIn[nI]) AND ((aIn[nI] - aIn[nI]) = (aIn[nI] - aIn[nI])); // 自反双判据（R79）/ the dual verdicts
    IF NOT bFin THEN // 非有限命中 / a non finite hit
        bError := TRUE; // 置故障（纪律②）/ raise the fault
        RETURN; // 早退（输出保持安全侧零）/ return early
    END_IF
END_FOR

// 段 4｜Hann 窗预加重与实部装填（虚部清零）/ segment 4, the Hann window and the loading
FOR nI := 0 TO nN - 1 DO // 逐点装填 / per point load
    IF bWinEn THEN // 加窗使能 / the window enabled
        aRe[nI] := aIn[nI] * (0.5 * (1.0 - COS(DL_FFT_TWOPI * DINT_TO_LREAL(nI) / DINT_TO_LREAL(nN - 1)))); // Hann 权重（nN ≥ 2 保证除子非零）/ the Hann weight, the divisor nonzero
    ELSE // 直通 / the pass through
        aRe[nI] := aIn[nI]; // 样本直通 / the sample direct
    END_IF
    aIm[nI] := 0.0; // 虚部清零 / clear the imaginary
END_FOR

// 段 5｜位反转序内排（CP 公开算法 ST 化）/ segment 5, the in place bit reversal
nJ := 0; // 反转索引清零 / clear the reversal index
FOR nI := 1 TO nN - 1 DO // 逐点重排 / per point reorder
    nBit := nN SHR 1; // 步进位起步 / start the stepping bit
    WHILE (nJ AND nBit) <> 0 DO // 逐位回退 / the bit rollback
        nJ := nJ - nBit; // 位清 / clear the bit
        nBit := nBit SHR 1; // 位右移 / shift the bit
    END_WHILE
    nJ := nJ + nBit; // 位置位 / set the bit
    IF nI < nJ THEN // 交换对（就地）/ the swap pair, in place
        fTr := aRe[nI];  aRe[nI] := aRe[nJ];  aRe[nJ] := fTr; // 实部交换 / swap the real
        fTi := aIm[nI];  aIm[nI] := aIm[nJ];  aIm[nJ] := fTi; // 虚部交换 / swap the imaginary
    END_IF
END_FOR

// 段 6｜基-2 蝶形主环（环长倍增有界终止，边界三）/ segment 6, the radix two butterfly main loop
nLen := 2; // 环长起步 / start the block length
WHILE nLen <= nN DO // 倍增推进 / the doubling advance
    nHalf := nLen SHR 1; // 环半长 / the half length
    fArg := -DL_FFT_TWOPI / DINT_TO_LREAL(nLen); // 基元旋转角（负向，正变换约定）/ the primitive angle, negative forward
    nBase := 0; // 环基址起步 / start the base
    WHILE nBase < nN DO // 环扫描 / the block scan
        FOR nJ := 0 TO nHalf - 1 DO // 半环内蝶形 / per butterfly in the half block
            fWr := COS(fArg * DINT_TO_LREAL(nJ)); // 旋转因子实部 / the twiddle real
            fWi := SIN(fArg * DINT_TO_LREAL(nJ)); // 旋转因子虚部 / the twiddle imaginary
            fTr := (aRe[nBase + nJ + nHalf] * fWr) - (aIm[nBase + nJ + nHalf] * fWi); // 上蝶实部 / the upper real
            fTi := (aRe[nBase + nJ + nHalf] * fWi) + (aIm[nBase + nJ + nHalf] * fWr); // 上蝶虚部 / the upper imaginary
            aRe[nBase + nJ + nHalf] := aRe[nBase + nJ] - fTr; // 下蝶写回 / the lower write back
            aIm[nBase + nJ + nHalf] := aIm[nBase + nJ] - fTi; // 下蝶写回 / the lower write back
            aRe[nBase + nJ] := aRe[nBase + nJ] + fTr; // 上蝶写回 / the upper write back
            aIm[nBase + nJ] := aIm[nBase + nJ] + fTi; // 上蝶写回 / the upper write back
        END_FOR
        nBase := nBase + nLen; // 环基址推进 / advance the base
    END_WHILE
    nLen := nLen + nLen; // 环长倍增（有界终止保证）/ double the block length, the bounded termination
END_WHILE
bValid := TRUE; // 变换完成 / the transform done
FC_DL_FftRadix2 := TRUE; // 受理 / accept
END_FUNCTION

(* ---- FC_DL_FilmSheetResistanceCalc.st ---- *)
(*
  DL Factory R88 | FC_DL_FilmSheetResistanceCalc
  功能：由电阻率与膜厚算方块电阻 Rs=ρ/t（厚度 nm 按 ÷1e7 换算 cm），并按带宽判合格
  开源溯源：无（clean-room 自研，依据公开工艺公式 方块电阻定义式 Rs=ρ/t，许可证=MIT，借鉴点=公式结构）
  规则：R1-R16 全遵守；R88 简单件标量形（纯标量入参出参，无循环体、无方法、无属性、无数组）
*)
FUNCTION FC_DL_FilmSheetResistanceCalc : REAL
VAR_INPUT
    fResistivityOhmCm : REAL := 1.0E-4; // 薄膜电阻率 ρ [Ω·cm] / film resistivity [ohm*cm]
    fThkNm : REAL := 500.0; // 薄膜厚度 t [nm] / film thickness [nm]
    fMinOhmSq : REAL := 0.1; // 方块电阻允许下限（工艺带宽） [Ω/□] / lower sheet resistance band [ohm/sq]
    fMaxOhmSq : REAL := 100.0; // 方块电阻允许上限（工艺带宽） [Ω/□] / upper sheet resistance band [ohm/sq]
END_VAR
VAR_OUTPUT
    fSheetOhmSq : REAL; // 方块电阻 Rs [Ω/□] / sheet resistance [ohm/sq]
    xInBand : BOOL; // TRUE=方块电阻落在允许带宽内 [-] / TRUE when inside the band [-]
END_VAR
VAR
    fThkCm : REAL; // 厚度换算为 cm（除零判据） [cm] / thickness in centimetres, the divisor [cm]
    fNmToCm : REAL; // nm→cm 换算因数 1e-7 [cm/nm] / conversion factor from nm to cm [cm/nm]
END_VAR

// 段 1｜出口预置
FC_DL_FilmSheetResistanceCalc := -1.0; // 哨兵返回 -1（无效） [-] / sentinel return -1, invalid [-]
fSheetOhmSq := 0.0; // 方块电阻预置零 [Ω/□] / sheet resistance preset zero [ohm/sq]
xInBand := FALSE; // 带宽位预置 FALSE（未判定前不认合格） [-] / band flag preset false [-]
fThkCm := 0.0; // 厚度 cm 值预置零 [cm] / thickness preset zero [cm]
fNmToCm := 0.0; // 换算因数预置零 [cm/nm] / conversion factor preset zero [cm/nm]

// 段 2｜非有限拦截 + 域闸
IF NOT (fResistivityOhmCm > -1.0E30 AND fResistivityOhmCm < 1.0E30) OR NOT (fThkNm > -1.0E30 AND fThkNm < 1.0E30) THEN
    RETURN; // 电阻率/膜厚任一非有限即拒算 [-] / any non finite input rejected [-]
END_IF
IF NOT (fMinOhmSq > -1.0E30 AND fMinOhmSq < 1.0E30) OR NOT (fMaxOhmSq > -1.0E30 AND fMaxOhmSq < 1.0E30) THEN
    RETURN; // 带宽上下限任一非有限则判据静默失效，故先拦 [Ω/□] / band limits must be finite [ohm/sq]
END_IF
IF fResistivityOhmCm < 1.0E-9 THEN
    RETURN; // 电阻率正域闸：须大于 1E-9（防零电阻率使结果恒零） [Ω·cm] / positive resistivity gate [ohm*cm]
END_IF
IF fThkNm < 1.0E-9 THEN
    RETURN; // 膜厚正域闸（同时是分母，防除零） [nm] / positive thickness, also the divisor [nm]
END_IF
IF fMinOhmSq <= 0.0 OR fMaxOhmSq <= fMinOhmSq THEN
    RETURN; // 带宽自洽闸：下限须为正、上限须严格大于下限 [Ω/□] / band consistency gate [ohm/sq]
END_IF

// 段 3｜计算
fNmToCm := 1.0E-7; // 1 nm = 1e-7 cm，换算因数装入 [cm/nm] / nm to cm factor [cm/nm]
fThkCm := fThkNm * fNmToCm; // nm × (cm/nm) = cm，厚度换算（等价 ÷1e7） [cm] / [nm] x [cm/nm] = [cm]
IF fThkCm < 1.0E-9 THEN
    RETURN; // 除法前分母闸：厚度 cm 值必须大于 1E-9 才可作除数 [cm] / denominator gate [cm]
END_IF
fSheetOhmSq := fResistivityOhmCm / fThkCm; // (Ω·cm) ÷ cm = Ω/□，方块电阻 [Ω/□] / [ohm*cm] / [cm] = [ohm/sq]

// 段 4｜判定与饱和
IF NOT (fSheetOhmSq > -1.0E30 AND fSheetOhmSq < 1.0E30) THEN
    RETURN; // 结果非有限再拦一次（防溢出成 Inf） [Ω/□] / re-check the result for finiteness [ohm/sq]
END_IF
xInBand := (fSheetOhmSq >= fMinOhmSq) AND (fSheetOhmSq <= fMaxOhmSq); // 双侧闭区间直比 [Ω/□] / closed two sided band compare [ohm/sq]

// 段 5｜出口自检
IF fSheetOhmSq < 0.0 THEN
    RETURN; // 出口自检：方块电阻不得为负（负值说明电阻率符号错） [Ω/□] / must not be negative [ohm/sq]
END_IF
FC_DL_FilmSheetResistanceCalc := fSheetOhmSq; // 返回方块电阻 [Ω/□] / return the sheet resistance [ohm/sq]
END_FUNCTION

(* ---- FC_DL_FixedFieldToInt.st ---- *)
(*==============================================================================
 * 组件名称 (Component)  : FC_DL_FixedFieldToInt
 * 溯源说明 (Provenance): 道莅 clean-room 防御性实现（IEC 61131-3 纯净实现，闭源文档仅借语义，零代码行）
 * 所属子库 (Sublibrary) : DL_MathData / DataFormat
 * 当前版本 (Version)    : 1.0.0
 * 兼容性   (Platform)   : CODESYS 3.5 / TwinCAT 3 / 汇川 InoProShop / 施耐德
 *                         Machine Expert；纯 IEC 61131-3（第 3 版），仅用
 *                         Standard.library 的 LEN / MID / MIN
 * 组件分类 (Category)   : 函数（FUNCTION）· 纯函数 · 定宽数值字段 → 整数
 * 功能一句话 (Summary)  : 把定宽十进制字段（前导零/空格填充、可选符号）解析成
 *                         DINT，非法字符精确报位置，超域给出饱和值并显式标记。
 *
 * 【填充与对齐规则（与 FC_DL_IntToFixedField 共用同一段口径原文）】
 *   ① 右对齐：数字永远贴字段右端，填充字符只在左侧。
 *   ② 填充字符为 '0' 或 ' '，剥离动作按 bAllowLeadingSpace 授权（零恒剥）。
 *   ③ 符号位占一位：零填充时符号贴最左（-0000042），空格填充时符号紧贴数字
 *      （     -42）——解析侧对两种排布等价，剥离填充后先取符号再取数字。
 *   ④ 宽度是契约：本件按 uWidth 与锁存串长的较小者参与解析，字段外的字符
 *      一律不看（定长报文的列位由此确定）。
 *
 * 本件存在的意义 (Why this unit exists)
 *   与 FC_DL_IntToFixedField 构成编码闭环。库内 FC_DL_StringToDint 解析「普通
 *   十进制串」，不看定宽列位、不剥零填充、不区分「非法字符」与「数值超域」，
 *   而 MES 回传的报文三者都需要：错字符要报第几位（现场改报文要定位），
 *   超域要能继续跑（饱和可观测），剥填充要留痕（口径可追）。
 *
 * 边界安全 (Boundary)
 *   ① uWidth < 1 → 故障 03AC；uWidth > 20 按物理上限 20 处理（码位表未分配该
 *      分支，不新开码，R90）；
 *   ② 剥填充后有效字符数为 0 → 故障 03AC（nErrPos 置 0，无单字符可指）；
 *   ③ 非数字字符 → 故障 03AB 且 nErrPos 精确到 1 基字符位，nValue 置 0；
 *   ④ 数值超 DINT 域 → 上界饱和 2147483647、下界饱和 −2147483647（哨兵值），
 *      置 bSaturated 与信息 045F，bValid 保持 TRUE——饱和是可观测的降级，
 *      与「非法字符」性质不同，后者 bValid 必须 FALSE；
 *   ⑤ 长度只取一次并锁存（R37/R38），其后所有上界都用该副本，绝不边解析边重算。
 * 遗留假设 (Assumption)
 *   累加升位到 LINT（R55①：取负前先升位复制到更宽类型）：LINT 可精确容纳
 *   −2147483648，故该值**可被本件精确解析**（不走哨兵路径），从而保证
 *   #1 → #2 的 round-trip 覆盖全 DINT 域；真正越界（> 2147483648）时下界
 *   饱和到 −2147483647 哨兵，bSaturated 为真，调用方须视为「不可用数值」。
 *   LINT 字面量 2147483648 依目标类型解释，属 P0 编译验证项（三平台各编译一次）。
 *
 * 错误码    : 16#0001_045E 已剥离前导填充（零或空格）——信息级，口径留痕
 *             16#0001_045F 数值超 DINT 域已饱和到边界值——信息级，饱和可观测
 *             16#0001_03AB 字段内出现非数字字符，nErrPos 给出首个非法位置——故障级
 *             16#0001_03AC 有效字符数为 0 或字段宽度非法——故障级
 *             16#0001_03AD 预留禁用（故障级，不得挪用）
 * 码位总账  : 16#0001_045E 用 / 16#0001_045F 用 ｜ 16#0001_03AB 用 / 16#0001_03AC 用 / 16#0001_03AD 预留
 * 状态机    : N/A —— 纯函数，两趟扫描（校验趟 + 累加趟），无顺序状态
 * 采样约定  : 纯组合函数，无定时器、无内部驻留状态
 * 依赖说明  : 无 DL_ 内部依赖；仅 Standard.library 的 LEN / MID / MIN
 * 验收向量  : V1 '00012345'/宽8 → 12345，uParsedLen=8，eErr=045E，TRUE
 *             V2 '     -42'/宽8 → -42，TRUE
 *             V3 '-2147483648'/宽11 → -2147483648（round-trip 主向量，不饱和）
 *             V4 '9999999999'/宽10 → 2147483647，bSaturated=TRUE，eErr=045F，TRUE
 *             V5 '00012X45'/宽8 → FALSE，nErrPos=6，nValue=0，eErr=03AB，bError=TRUE
 *             V6 '        '/宽8 → FALSE，eErr=03AC
 *             V7 宽 0 → FALSE，eErr=03AC，nErrPos=0
 * 红线自检  : 全局变量声明零使用 / 外部变量访问零使用 / 物理地址零使用 ｜ 纯 IEC 61131-3 ｜ 零浮点
 *             比较、零除法 ｜ 循环全部带 nGuard ｜ 数组写入前置界检 ｜ 全变量
 *             双语同行注释 ｜ 状态机 N/A ｜ 无定时器实例 ｜ 无魔法数
 * 修订历史  : 2026-11-16  v1.0.0  首版入库（R22 · 批 1 · 定宽数值字段族）
 *============================================================================*)

FUNCTION FC_DL_FixedFieldToInt : BOOL
VAR_INPUT
    sField             : STRING(20);           // 待解析定宽字段 [ASCII] / fixed width field to parse [ASCII]
    uWidth             : UINT := 8;            // 参与解析的字符数 [字符]，范围 1~20 / characters to parse [char], range 1~20
    bAllowLeadingSpace : BOOL := TRUE;         // 是否允许剥离前导空格（零恒剥） / allow stripping leading spaces, zeros always stripped
    bAllowSign         : BOOL := TRUE;         // 是否接受前置 '+'/'-' 号 / accept a leading plus or minus sign
END_VAR
VAR_OUTPUT
    nValue      : DINT;                        // 解析结果，超域时取饱和值 [无量纲] / parsed value, saturated when out of range
    uParsedLen  : UINT;                        // 成功解析的数字位数 [位] / number of digits parsed
    nErrPos     : UINT;                        // 1 基首个非法字符位置，0 表示无 [位置] / 1-based first illegal position, 0 means none
    bSaturated  : BOOL;                        // 数值超 DINT 域已饱和标志 / value saturated at the DINT boundary
    eErr        : UDINT;                       // 错误码，0 表示无错 / error code, 0 means no error
    bError      : BOOL;                        // 故障级标志，仅故障级错误置位 / fault-class flag, set only on fault-level codes
    bValid      : BOOL;                        // 结果可用标志（饱和时仍为 TRUE） / result usable flag, still TRUE when saturated
END_VAR
VAR
    nLenLock    : INT;                         // 锁存的字段长度 [字符]，全件唯一长度源 / latched field length, the single length source
    nLenRaw     : INT;                         // LEN 的原始读数 [字符] / raw LEN reading
    nWUse       : INT;                         // 生效解析宽度 [字符] / effective parse width
    nParseLen   : INT;                         // 实际参与解析的字符数 [字符] / characters actually parsed
    nPos        : INT;                         // 当前扫描位置，1 基 [位置] / current scan position, 1-based
    nDigitCount : INT;                         // 已采集数字位个数 [位] / collected digit count
    nI          : INT;                         // 数字位遍历下标 [索引] / digit index
    nGuard      : INT;                         // 循环守卫计数器 [次] / loop guard counter
    nDigitV     : INT;                         // 单字符对应的数值 0~9 [无量纲] / numeric value of a single character
    nScanV      : INT;                         // 查表扫描下标 0~9 [索引] / table scan index
    bNegSign    : BOOL;                        // 字段带负号 / field carries a minus sign
    bStripped   : BOOL;                        // 发生过剥填充动作 / padding was stripped
    bStopStrip  : BOOL;                        // 剥离循环终止标志 / strip loop stop flag
    bIsDigit    : BOOL;                        // 当前字符是否数字 / current character is a digit
    sCh         : STRING(1);                   // 当前字符 [ASCII] / current character
    aDig        : ARRAY[1..20] OF USINT;       // 数字位缓存，1 基 [无量纲] / digit cache, 1-based
    liAcc       : LINT;                        // 升位累加器，防 DINT 回绕 [无量纲] / widened accumulator, avoids DINT wrap
END_VAR
VAR CONSTANT
    DL_FIELD_MAX   : UINT := 20;               // STRING(20) 物理上限 [字符]，禁写成 255 / physical bound of STRING(20), never 255
    DL_W_MIN_U     : UINT := 1;                // 宽度下限的无符号副本 [字符] / unsigned copy of the width lower bound
    DL_W_MAX       : INT := 20;                // 宽度上限 [字符] / width upper bound
    DL_DIGIT_MAX   : INT := 20;                // 字段内最多数字位 [位]，等于串上限 / maximum digits inside the field
    DL_DINT_DIGITS : INT := 10;                // DINT 十进制最大位数 [位]，超过即必饱和 / DINT maximum decimal digits
    DL_GUARD_MAX   : INT := 24;                // 循环守卫上限 [次]，大于串上限即安全 / loop guard, larger than the field
    DL_TEN         : LINT := 10;               // 十进制基数 [无量纲] / decimal radix
    DL_POS_ONE     : INT := 1;                 // 单字符长度与位置基数 [字符] / single-char length and position base
    DL_DIGITS      : STRING(10) := '0123456789'; // 数字字符表，字符→数值靠查表 / digit table, character to value by lookup
    DL_PAD_ZERO    : STRING(1) := '0';         // 零填充字符 [字符] / zero pad character
    DL_PAD_SPACE   : STRING(1) := ' ';         // 空格填充字符 [字符] / space pad character
    DL_SIGN_PLUS   : STRING(1) := '+';         // 正号字符 [字符] / plus sign character
    DL_SIGN_MINUS  : STRING(1) := '-';         // 负号字符 [字符] / minus sign character
    DL_LINT_MAX    : LINT := 2147483647;       // DINT 上界 [无量纲] / DINT upper bound
    DL_LINT_MIN_ABS: LINT := 2147483648;       // DINT 下界绝对值 [无量纲] / absolute value of the DINT lower bound
    DL_DINT_MAX    : DINT := 2147483647;       // DINT 上界饱和值 [无量纲] / DINT upper saturation value
    DL_DINT_MIN_SAT: DINT := -2147483647;      // DINT 下界哨兵饱和值 [无量纲] / DINT lower sentinel saturation value
    DL_DIG_LAST    : INT := 9;                 // 数字表末位下标 [索引] / last index of the digit table
END_VAR

(*------------------------------------------------------------------------------
 * 段 1｜返回值与输出预置（L1/L9：任何失败出口都不留脏值）
 *      Preset the return value and every output, no stale value on any exit
 *-----------------------------------------------------------------------------*)
FC_DL_FixedFieldToInt := FALSE;                // 返回值预置失败 / preset to FALSE
nValue      := 0;                              // 结果预置 0 [无量纲] / result preset to zero
uParsedLen  := 0;                              // 解析位数预置 0 [位] / parsed length preset to zero
nErrPos     := 0;                              // 非法位置预置 0（无） / illegal position preset to none
bSaturated  := FALSE;                          // 饱和标志预置 FALSE / saturation flag preset to FALSE
eErr        := 16#0000_0000;                   // 错误码预置无错 / error code preset to none
bError      := FALSE;                          // 故障标志预置 FALSE / fault flag preset to FALSE
bValid      := FALSE;                          // 结果可用预置 FALSE / usable flag preset to FALSE
nLenLock    := 0;                              // 锁存长度预置 0 / latched length preset to zero
nWUse       := DL_W_MAX;                       // 生效宽度预置上限 / effective width preset to the upper bound
nParseLen   := 0;                              // 参与解析字符数预置 0 / parsed character count preset to zero
nPos        := DL_POS_ONE;                     // 扫描位置从 1 起 / scan starts at position one
nDigitCount := 0;                              // 数字位个数预置 0 / digit count preset to zero
nGuard      := 0;                              // 守卫预置 0 / guard preset to zero
bNegSign    := FALSE;                          // 负号标志预置 FALSE / negative flag preset to FALSE
bStripped   := FALSE;                          // 剥填充标志预置 FALSE / strip flag preset to FALSE
bStopStrip  := FALSE;                          // 剥离终止标志预置 FALSE / strip stop flag preset to FALSE
liAcc       := 0;                              // 累加器预置 0 / accumulator preset to zero

(*------------------------------------------------------------------------------
 * 段 2｜字段宽度闸门（宽度非法属故障级；超物理上限按上限处理不留码）
 *      Width gate: an illegal width latches a fault, the physical ceiling is clamped
 *-----------------------------------------------------------------------------*)
IF uWidth < DL_W_MIN_U THEN
    eErr    := 16#0001_03AC;                   // 故障级：宽度非法 / fault: illegal width
    bError  := TRUE;                           // 置故障标志 / raise the fault flag
    bValid  := FALSE;                          // 结果不可用 / result unusable
    nErrPos := 0;                              // 无单字符可指 / no specific character to point at
    RETURN;                                    // 统一后处理已在本段完成 / the exit is fully post-processed here
ELSIF uWidth > DL_FIELD_MAX THEN
    nWUse := DL_W_MAX;                         // 超物理上限按 20 处理（不新开码，R90） / clamped to the physical ceiling, no new code
ELSE
    nWUse := UINT_TO_INT(uWidth);              // 域内直通 / passed through inside the domain
END_IF

(*------------------------------------------------------------------------------
 * 段 3｜长度只取一次并锁存（R37/R38：绝不边解析边重算）
 *      Latch the length exactly once, never recompute it while parsing
 *-----------------------------------------------------------------------------*)
nLenRaw := LEN(sField);                        // 唯一一次取长度 / the single length read
IF nLenRaw < 0 THEN
    nLenRaw := 0;                              // 结构性兜底：LEN 不应为负 / structural fallback, LEN should never be negative
END_IF
nLenLock := nLenRaw;                           // 锁存副本，其后全部比较都用它 / latched copy used by every later comparison
nParseLen := MIN(nWUse, nLenLock);             // 实际解析长度 = 宽度与串长的较小者 / the smaller of width and length
IF nParseLen < 0 THEN
    nParseLen := 0;                            // 结构性兜底 / structural fallback
END_IF

(*------------------------------------------------------------------------------
 * 段 4｜剥离前导填充（零恒剥，空格按授权剥；剥过即留痕 045E）
 *      Strip leading padding, zeros always, spaces only when allowed
 *-----------------------------------------------------------------------------*)
WHILE (NOT bStopStrip) AND (nPos <= nParseLen) AND (nGuard <= DL_GUARD_MAX) DO
    sCh := MID(sField, DL_POS_ONE, nPos);      // 取当前字符 [ASCII] / read the current character
    IF sCh = DL_PAD_ZERO THEN
        nPos      := nPos + DL_POS_ONE;        // 前导零：跳过 / leading zero skipped
        bStripped := TRUE;                     // 剥填充留痕 / padding stripped, recorded
    ELSIF bAllowLeadingSpace AND (sCh = DL_PAD_SPACE) THEN
        nPos      := nPos + DL_POS_ONE;        // 授权的前导空格：跳过 / authorised leading space skipped
        bStripped := TRUE;                     // 剥填充留痕 / padding stripped, recorded
    ELSE
        bStopStrip := TRUE;                    // 遇到非填充字符即停 / stop at the first non-pad character
    END_IF
    nGuard := nGuard + DL_POS_ONE;             // 守卫累计，防死循环 / guard incremented, prevents a dead loop
END_WHILE

(*------------------------------------------------------------------------------
 * 段 5｜符号位（授权才接受；不授权则按非法字符定位）
 *      Sign position, accepted only when authorised, otherwise reported as illegal
 *-----------------------------------------------------------------------------*)
IF nPos <= nParseLen THEN
    sCh := MID(sField, DL_POS_ONE, nPos);      // 取候选符号字符 / read the candidate sign character
    IF (sCh = DL_SIGN_MINUS) OR (sCh = DL_SIGN_PLUS) THEN
        IF bAllowSign THEN
            bNegSign := (sCh = DL_SIGN_MINUS); // 负号判据（字符比较，非浮点） / negative test, a character comparison
            nPos     := nPos + DL_POS_ONE;     // 符号位已消费 / the sign position is consumed
        ELSE
            eErr    := 16#0001_03AB;           // 故障级：不允许符号却出现符号 / fault: a sign appeared although not allowed
            bError  := TRUE;                   // 置故障标志 / raise the fault flag
            bValid  := FALSE;                  // 结果不可用 / result unusable
            nErrPos := INT_TO_UINT(nPos);      // 非法位置精确到字符 / illegal position pinpointed
            nValue  := 0;                      // 结果归零 / result zeroed
            RETURN;                            // 统一后处理完成 / exit fully post-processed
        END_IF
    END_IF
END_IF

(*------------------------------------------------------------------------------
 * 段 6｜校验趟：逐字符判数字并缓存数值，首个非法字符即定位（不早退留脏值）
 *      Validation pass: every character must be a digit, the first illegal one is located
 *-----------------------------------------------------------------------------*)
WHILE (nPos <= nParseLen) AND (nGuard <= (DL_GUARD_MAX * 2)) DO
    sCh      := MID(sField, DL_POS_ONE, nPos); // 取当前字符 / read the current character
    bIsDigit := FALSE;                         // 数字判据预置 FALSE / digit test preset to FALSE
    nDigitV  := 0;                             // 数值预置 0 / numeric value preset to zero
    nScanV   := 0;                             // 查表下标预置 0 / table index preset to zero
    WHILE (nScanV <= DL_DIG_LAST) AND (NOT bIsDigit) DO
        IF sCh = MID(DL_DIGITS, DL_POS_ONE, nScanV + DL_POS_ONE) THEN
            bIsDigit := TRUE;                  // 命中数字表 / a table entry matched
            nDigitV  := nScanV;                // 下标即数值 / the index is the numeric value
        ELSE
            nScanV := nScanV + DL_POS_ONE;     // 继续查下一位 / advance to the next table entry
        END_IF
    END_WHILE

    IF NOT bIsDigit THEN
        eErr    := 16#0001_03AB;               // 故障级：非数字字符 / fault: non-digit character
        bError  := TRUE;                       // 置故障标志 / raise the fault flag
        bValid  := FALSE;                      // 结果不可用 / result unusable
        nErrPos := INT_TO_UINT(nPos);          // 1 基位置精确到字符 / 1-based position pinpointed
        nValue  := 0;                          // 结果归零，绝不交出半解析值 / result zeroed, no half-parsed value
        uParsedLen := 0;                       // 解析位数归零 / parsed length zeroed
        RETURN;                                // 统一后处理完成 / exit fully post-processed
    END_IF

    IF (nDigitCount + DL_POS_ONE) <= DL_DIGIT_MAX THEN
        aDig[nDigitCount + DL_POS_ONE] := INT_TO_USINT(nDigitV); // 缓存数字（前置界检） / cache the digit after a bounds check
        nDigitCount := nDigitCount + DL_POS_ONE;                 // 位数累计 / digit count incremented
    END_IF
    nPos   := nPos + DL_POS_ONE;               // 位置推进 / position advanced
    nGuard := nGuard + DL_POS_ONE;             // 守卫累计 / guard incremented
END_WHILE

(*------------------------------------------------------------------------------
 * 段 7｜有效字符数为 0 的判定（全填充字段不是 0，是「没有数字」）
 *      Zero effective characters: an all-pad field carries no number at all
 *-----------------------------------------------------------------------------*)
IF nDigitCount = 0 THEN
    eErr    := 16#0001_03AC;                   // 故障级：有效字符数为 0 / fault: zero effective characters
    bError  := TRUE;                           // 置故障标志 / raise the fault flag
    bValid  := FALSE;                          // 结果不可用 / result unusable
    nErrPos := 0;                              // 无单字符可指 / no specific character to point at
    nValue  := 0;                              // 结果归零 / result zeroed
    RETURN;
END_IF

(*------------------------------------------------------------------------------
 * 段 8｜累加趟：位数超 DINT 位宽必饱和（先判位宽，绝不进累加，杜绝 LINT 溢出）
 *      Accumulation: more than ten digits saturates immediately, so LINT never overflows
 *-----------------------------------------------------------------------------*)
IF nDigitCount > DL_DINT_DIGITS THEN
    IF bNegSign THEN
        nValue := DL_DINT_MIN_SAT;             // 下界哨兵值（−2147483648 留给精确路径） / lower sentinel, the exact value has its own path
    ELSE
        nValue := DL_DINT_MAX;                 // 上界饱和 / saturated at the upper bound
    END_IF
    bSaturated := TRUE;                        // 饱和可观测 / saturation made observable
    eErr       := 16#0001_045F;                // 信息级：已饱和（优先于 045E） / informational: saturated, takes precedence over 045E
    uParsedLen := INT_TO_UINT(nDigitCount);    // 解析位数仍如实上报 / parsed length still reported truthfully
    bValid     := TRUE;                        // 饱和是可观测降级，结果仍可用 / degraded but observable, still usable
    FC_DL_FixedFieldToInt := TRUE;             // 返回成功 / return success
    RETURN;
END_IF

liAcc := 0;                                    // 累加器清零 / accumulator cleared
FOR nI := DL_POS_ONE TO nDigitCount DO
    liAcc := liAcc * DL_TEN + INT_TO_LINT(aDig[nI]); // 升位累加，LINT 内无回绕 / widened accumulation, no wrap inside LINT
END_FOR

(*------------------------------------------------------------------------------
 * 段 9｜边界仲裁与出口（精确路径覆盖 −2147483648，越界才走哨兵）
 *      Boundary arbitration: the exact path covers -2147483648, only true overflow saturates
 *-----------------------------------------------------------------------------*)
IF bNegSign THEN
    IF liAcc > DL_LINT_MIN_ABS THEN
        nValue     := DL_DINT_MIN_SAT;         // 真越界：下界哨兵 / true overflow, lower sentinel
        bSaturated := TRUE;                    // 饱和可观测 / saturation observable
        eErr       := 16#0001_045F;            // 信息级：已饱和 / informational: saturated
    ELSE
        nValue := LINT_TO_DINT(-liAcc);        // 精确负值（含 −2147483648） / exact negative value, including the DINT minimum
    END_IF
ELSE
    IF liAcc > DL_LINT_MAX THEN
        nValue     := DL_DINT_MAX;             // 上界饱和 / saturated at the upper bound
        bSaturated := TRUE;                    // 饱和可观测 / saturation observable
        eErr       := 16#0001_045F;            // 信息级：已饱和 / informational: saturated
    ELSE
        nValue := LINT_TO_DINT(liAcc);         // 精确正值 / exact positive value
    END_IF
END_IF

(*------------------------------------------------------------------------------
 * 段 10｜码位优先级与出口（饱和码优先于剥填充码，信息级不置 bError）
 *      Code precedence and exit: saturation outranks stripping, info codes never raise bError
 *-----------------------------------------------------------------------------*)
IF bStripped AND (eErr = 16#0000_0000) THEN
    eErr := 16#0001_045E;                      // 信息级：已剥离前导填充 / informational: leading padding stripped
END_IF

uParsedLen := INT_TO_UINT(nDigitCount);        // 解析位数出口 [位] / parsed length outlet
bValid     := TRUE;                            // 结果可用 / result usable
FC_DL_FixedFieldToInt := TRUE;                 // 解析成功 / parse succeeded
END_FUNCTION

(* ---- FC_DL_FloorEx.st ---- *)
(*
    FC_DL_FloorEx —— 向下取整防御包装（向 -∞，DINT 范围钳位 + NaN 拦截）
    ------------------------------------------------------------------
    分类      : DL_MathData / Math-Round
    前缀      : FC_DL_
    版本      : 1.0.0
    溯源      : IEC 61131-3 标准语义的道莅防御性实现
                （内部委托平台内建函数，外围统一错误码/钳位/双语文档；
                  未复制任何闭源厂商源码，参考实现仅限 MIT/Apache 许可）
    平台      : 纯 IEC 61131-3，CODESYS / TwinCAT / InoProShop 通用
    作者      : 道莅代码库 · PLC编程专家（R15）
    ------------------------------------------------------------------
    功能说明  : 向负无穷方向取整（委托内建 FLOOR），负小数如 -1.2 得
                -2。NaN 输入拦截返回 0 并置 16#0001_0190；先以 LREAL 承载 FLOOR
                结果再做 DINT 范围闸（FLOOR 本身不会上溢 LREAL），超
                [-2147483648, 2147483647] 时钳位到边界并置 16#0001_025E，bValid=
                FALSE；无穷输入被范围闸自然拦截。范围内再经 LREAL_TO_DINT
                显式转换，转换永不溢出。
    错误码    : 0000 正常 / 16#0001_0190 入参越界（NaN 已归零） / 16#0001_025E 上溢下溢（已钳位到 DINT 边界）
    修订记录  : 2026-11-16 v1.0.0 首次入库（R15）
*)
FUNCTION FC_DL_FloorEx : DINT
VAR_INPUT
    lrIn : LREAL; // 输入实数 [无量纲]，任意有限值或 NaN/无穷 / input real value [dimensionless], any finite value or NaN/inf
END_VAR
VAR_OUTPUT
    eErr : UDINT; // 错误码，0=正常，1=入参越界，2=上溢下溢 / error id, 0=ok, 1=input out of domain, 2=overflow or underflow
    bError   : BOOL; // 是否出错，eErr 非 0 时为 TRUE / error flag, TRUE when eErr is nonzero
    bValid   : BOOL; // 输出是否有效可用，钳位降级时为 FALSE / output valid, FALSE for clamped degraded results
END_VAR
VAR
    lrR : LREAL; // FLOOR 结果中间量 [无量纲]，LREAL 承载不溢出 / intermediate FLOOR result [dimensionless], carried in LREAL without overflow
END_VAR
VAR CONSTANT
    DL_FL_HI : LREAL := 2147483647.0; // DINT 上界 [无量纲]，超过即钳位 / DINT upper bound [dimensionless], beyond clamped
    DL_FL_LO : LREAL := -2147483648.0; // DINT 下界 [无量纲]，低于即钳位 / DINT lower bound [dimensionless], below clamped
END_VAR

// 段 1｜返回值与错误状态预置，任何早退路径不留脏码 / segment 1, preset return value and error states
FC_DL_FloorEx := 0; // 返回值预置安全值 0 / preset return to safe value 0
eErr      := 16#0000_0000; // 错误码预置正常 / preset error id to ok
bError        := FALSE; // 错误标志预置无错 / preset error flag to FALSE
bValid        := TRUE; // 有效标志预置可用 / preset valid flag to TRUE

// 段 2｜NaN 拦截：自不等判据，归零早退，不进内核 / segment 2, NaN interception by self-inequality, zeroed early exit
IF lrIn <> lrIn THEN
    eErr := 16#0001_0190; // 信息级：输入 NaN，已归零 / informational, NaN input, zeroed
    bError   := TRUE; // 置错误标志 / raise error flag
    bValid   := FALSE; // 输出不可用 / output invalid
    RETURN; // 返回预置安全值 0 / return preset safe value 0
END_IF

// 段 3｜委托内建 FLOOR（向 -∞ 取整），LREAL 承载结果，无穷输入得无穷 / segment 3, delegation to built-in FLOOR toward minus infinity, LREAL carry, infinite input stays infinite
lrR := FLOOR(lrIn); // 委托内建 FLOOR 内核，不自实现取整内核 / delegate to built-in FLOOR kernel

// 段 4｜DINT 范围闸：超界钳位并置 16#0001_025E（无穷输入在此被拦截） / segment 4, DINT range gate, clamp beyond bounds with code 2, infinite input intercepted here
IF lrR > DL_FL_HI THEN
    FC_DL_FloorEx := 2147483647; // 上溢钳位到 DINT 上界 / overflow clamped to the DINT upper bound
    eErr      := 16#0001_025E; // 上溢码 / overflow code
    bError        := TRUE; // 置错误标志 / raise error flag
    bValid        := FALSE; // 钳位值非真实取整 / clamped value is not the true floor
    RETURN;
ELSIF lrR < DL_FL_LO THEN
    FC_DL_FloorEx := -2147483648; // 下溢钳位到 DINT 下界 / underflow clamped to the DINT lower bound
    eErr      := 16#0001_025E; // 下溢码 / underflow code
    bError        := TRUE; // 置错误标志 / raise error flag
    bValid        := FALSE; // 钳位值非真实取整 / clamped value is not the true floor
    RETURN;
END_IF

// 段 5｜范围内显式转换输出（转换永不溢出） / segment 5, explicit in-range conversion and output
FC_DL_FloorEx := LREAL_TO_DINT(lrR); // 范围内显式转换 / explicit in-range conversion
END_FUNCTION

(* ---- FC_DL_FloorToMultipleInt.st ---- *)
(*==============================================================================
 * 组件名称 : FC_DL_FloorToMultipleInt ｜ 子库 : DL_MathData ｜ v1.0.0 ｜ 2026-11-23
 * 平台     : CODESYS 3.5 / TwinCAT 3 / InoProShop / Machine Expert（纯 IEC，无厂商库）
 * 功能简介 : 整数向下（朝 -∞ 方向）对齐到 nMultiple 的倍数。纯整数算术
 *            实现：整除截取得基准，仅当值小于基准时退位一个倍数；
 *            退位前做 DINT 下限反算防饱和溢出，越限饱和到 -2147483648。
 * 契约     : 返回向下对齐结果；nMultiple <= 0 恒返回 0；
 *            纯函数无状态、同输入同输出。
 * 依赖     : 无 DL_ 内部依赖（本批自足实现）
 * 红线自检 : R1 零全局 R2 零%I/%Q R3 纯IEC R4 非法倍数返 0 + 下限反算防溢出
 *            R5 双语注释 R6 N/A（无状态机） R7 N/A（无定时器实例）
 * 修订历史 : 2026-11-23 R78-B1 对齐取整族模板派生首版
 *============================================================================*)
FUNCTION FC_DL_FloorToMultipleInt : DINT
VAR_INPUT
    nValue : DINT;          // 输入整数 / Input integer value
    nMultiple : DINT;       // 对齐倍数，须 > 0 / Alignment multiple, must be > 0
END_VAR
VAR
    nLo : DINT;             // 向零截断的基准倍数值 / Truncated-toward-zero base multiple
END_VAR
IF nMultiple <= 0 THEN
    FC_DL_FloorToMultipleInt := 0;      // 非法倍数返 0 / Invalid multiple returns 0
    RETURN;
END_IF
nLo := (nValue / nMultiple) * nMultiple;    // 整除截取得基准 / Base via integer division truncation
IF nValue < nLo THEN
    IF nLo >= (-2147483648 + nMultiple) THEN
        nLo := nLo - nMultiple;             // 向 -∞ 对齐到下一倍数 / Align down to next multiple
    ELSE
        nLo := -2147483648;                 // 退位将溢出，饱和到 DINT 下限 / Saturation at DINT min
    END_IF
END_IF
FC_DL_FloorToMultipleInt := nLo;            // 输出向下对齐结果 / Output floor-aligned result
END_FUNCTION

(* ---- FC_DL_FuelCellStoichAirCalc.st ---- *)
(*
  DL Factory R88 | FC_DL_FuelCellStoichAirCalc
  功能：算燃料电池空气计量比 λ=实际空气质量流量/理论需求量（理论=O2 摩尔流×M_O2/0.232），λ<1.5 判偏稀
  开源溯源：无（clean-room 自研，依据公开工艺公式 电化学氧耗与空气计量比定义式 λ=m_air/m_air,st，许可证=MIT，借鉴点=公式结构）
  规则：R1-R16 全遵守；R88 简单件标量形（纯标量入参出参，无循环体、无方法、无属性、无数组）
*)
FUNCTION FC_DL_FuelCellStoichAirCalc : REAL
VAR_INPUT
    fCurrentA : REAL := 300.0; // 电堆电流 I [A] / stack current [A]
    fCells : REAL := 400.0; // 串联单胞数量 n [个] / number of series cells [-]
    fAirFlowKgH : REAL := 60.0; // 实测干空气质量流量 [kg/h] / measured dry air mass flow [kg/h]
    fLambdaMin : REAL := 1.5; // 计量比合格下限（λ<1.5 判偏稀） [-] / lean threshold [-]
END_VAR
VAR_OUTPUT
    fLambda : REAL; // 空气计量比 λ [-] / air stoichiometry [-]
    xLean : BOOL; // TRUE=计量比低于下限，偏稀需加风 [-] / TRUE when the air is lean [-]
END_VAR
VAR
    fFaradayC : REAL; // 法拉第常数 F [C/mol] / faraday constant [C/mol]
    fFourF : REAL; // 分母 4F（每摩 O2 需 4 mol 电子） [C/mol] / the 4F divisor [C/mol]
    fAirTheoKgH : REAL; // 理论干空气质量流量（除零判据） [kg/h] / theoretical air flow, the divisor [kg/h]
END_VAR

// 段 1｜出口预置
FC_DL_FuelCellStoichAirCalc := -1.0; // 哨兵返回 -1（无效） [-] / sentinel return -1, invalid [-]
fLambda := 0.0; // 计量比预置零 [-] / stoichiometry preset zero [-]
xLean := FALSE; // 偏稀位预置 FALSE（未判定前不报警） [-] / lean flag preset false [-]

// 段 2｜非有限拦截 + 域闸
IF NOT (fCurrentA > -1.0E30 AND fCurrentA < 1.0E30) OR NOT (fCells > -1.0E30 AND fCells < 1.0E30) THEN
    RETURN; // 电流/单胞数任一非有限即拒算 [-] / any non finite input rejected [-]
END_IF
IF NOT (fAirFlowKgH > -1.0E30 AND fAirFlowKgH < 1.0E30) OR NOT (fLambdaMin > -1.0E30 AND fLambdaMin < 1.0E30) THEN
    RETURN; // 空气流量/下限任一非有限则判据静默失效，故先拦 [-] / these pins must be finite [-]
END_IF
IF fCurrentA < 0.0 OR fCells < 1.0 OR fAirFlowKgH < 0.0 THEN
    RETURN; // 电流非负闸 + 单胞下限闸 + 空气流量非负闸 [A, 个, kg/h] / non negative gates
END_IF
IF fLambdaMin <= 0.0 THEN
    RETURN; // 下限正域闸：非正下限会使判据恒假 [-] / positive threshold gate [-]
END_IF

// 段 3｜计算（I→O2 mol/s→空气质量→kg/h 链路，逐项量纲见行尾注释）
fFaradayC := 96485.0; // 法拉第常数装入 [C/mol] / load the faraday constant [C/mol]
fFourF := 4.0 * fFaradayC; // 4 × C/mol = C/mol，每摩 O2 需 4 摩电子 [C/mol] / [C/mol]
IF fFourF < 1.0E-9 THEN
    RETURN; // 除法前分母闸：4F 必须大于 1E-9 才可作除数 [C/mol] / denominator gate [C/mol]
END_IF
fAirTheoKgH := (fCurrentA * fCells / fFourF) * 32.0 * 0.001 / 0.232 * 3600.0; // (mol/s)×32 g/mol×0.001 kg/g÷0.232(空气质量分数)×3600 s/h = kg/h [kg/h] / [kg/h]
IF fAirTheoKgH < 1.0E-9 THEN
    RETURN; // 除法前分母闸：理论空气量必须大于 1E-9（零电流时无意义） [kg/h] / denominator gate [kg/h]
END_IF
fLambda := fAirFlowKgH / fAirTheoKgH; // (kg/h) ÷ (kg/h) = 无量纲，计量比 λ [-] / dimensionless stoichiometry [-]

// 段 4｜判定与饱和
IF NOT (fLambda > -1.0E30 AND fLambda < 1.0E30) THEN
    RETURN; // 结果非有限再拦一次 [-] / re-check the result for finiteness [-]
END_IF
xLean := fLambda < fLambdaMin; // 严格小于下限判偏稀，等于下限仍判合格 [-] / strict compare against the threshold [-]

// 段 5｜出口自检
IF fLambda < 1.0 THEN
    xLean := TRUE; // 出口自检：λ<1 已属缺氧区（低于电化学计量），强制置偏稀 [-] / below unity is oxygen starved [-]
END_IF
FC_DL_FuelCellStoichAirCalc := fLambda; // 返回空气计量比 λ [-] / return the air stoichiometry [-]
END_FUNCTION

(* ---- FC_DL_GcdUdintCalc.st ---- *)
(*
  ==================================================================
  组件名 Component  : FC_DL_GcdUdintCalc
  分类   Category   : DL_MathData
  前缀   Naming     : FC_DL_ ｜ b/n/u/f/t/e/st 类型前缀制（R265）
  码位   Code ID    : 16#0001_0663（信息级）｜ 16#0001_0664（故障级）
  版本   Version    : 1.0.0
  复杂度 Complexity  : 低
  功能   Purpose    : UDINT 最大公约数（欧几里得迭代 + WHILE 守卫计数），供
                      电子齿轮比约分、脉冲当量配比、采样周期同步等调用方；
                      返回 GCD(nA, nB)，双零入参返回 0 哨兵 + 信息级。
  开源溯源 Origin    : T0 数论原子补口（内部来源，零检索）；欧几里得算法为
                      公共领域数学事实；WHILE 守卫计数为道莅防御性范式。
  许可证 License    : MIT
  参考   Reference  : IEC 61131-3:2013 §6.6.4 WHILE / MOD 语义；欧几里得
                      算法（公共领域数学事实）
  平台   Platform   : 纯 IEC 61131-3（WHILE / MOD / 比较），三平台通用
  依赖   Depends    : 无（零委托、零库件）
  分工声明 Split     : FC_DL_IntLcmSafeUdint（最小公倍数，R79 入库，委托本件 GCD 作除子；原头注写的 FC_DL_LcmUdintCalc 为规划期名，实际入库名以本行为准）
                      为互补件（互引）；本件只算 GCD，不做 LCM（LCM 含
                      乘法溢出域，职责分离，R216）。
  归属 Ownership     : 本件无 TYPE 声明；全部引脚为 IEC 标准原生类型。
  ------------------------------------------------------------------
  边界 Boundary     :
                      一 双零哨兵（nA = 0 且 nB = 0）：GCD 数学上无定义，
                         返回 0 哨兵 + 信息级 0663 + bValid = TRUE（调用方
                         以 0 值即可甄别，不置 bError——组态缺省不是运行
                         故障）；单零入参按 GCD(x, 0) = x 口径返回非零方；
                      二 MOD 除零防：循环条件 nY <> 0 已证除子非零，除法段
                         不可达（R1 教训出厂即正确）；
                      三 WHILE 守卫计数（DL_GCD_GUARDMAX = 64）：纯 IEC 语义
                         下欧几里得迭代余量单调递减、必在极小步数内终止，
                         守卫理论不可达；触发路径仅为平台 UDINT MOD 异常
                         回绕类非标行为（安全断言反例声明）；守卫命中 →
                         故障级 0664 + 返回 0 哨兵 + bValid = FALSE；
                      四 迭代计数 nIter 外显 [次]，供调用方审计收敛步数；
                      五 纯函数：无记忆量、无定时器、无边沿实例，每调用重算；
                      六 无全局、无外部变量、无物理地址。
  错误码 Codes      :
    16#0001_0663【信息级】双零入参（GCD 无定义，返回 0 哨兵，不置 bError）
    16#0001_0664【故障级】WHILE 守卫计数越限（平台异常回绕类，理论不可达防御）
  码位反证 Note     :
    0663 与 0664 不可合并：0663 出口 bValid = TRUE（哨兵 0 是合法甄别结果），
    0664 出口 bValid = FALSE（结果不可用），bValid 可唯一区分两场景，按 R90
    分立；单零入参（GCD(x, 0) = x）为正常数学口径，无码。
  验收 Acceptance   :
    算法已证（脚本）：未跑 ｜ 编译器已证（三平台）：未跑
    V1 GCD(48, 36) = 12；V2 GCD(17, 5) = 1（互质）
    V3 GCD(7, 0) = 7 / GCD(0, 7) = 7（单零口径）
    V4 GCD(0, 0) → 0 哨兵 + 信息级 0663（bError = FALSE）
    V5 nIter 审计：V1 场景 nIter = 2（48,36 → 36,12 → 12,0）
    V6 守卫命中（强改平台异常注入）→ 码 0664 + bValid = FALSE + 返回 0
  修订记录 Revision  :
    2026-11-21  v1.0.0  R64 首版（批 1 · 序号 3，T0 数论原子补口）
  ==================================================================
*)
FUNCTION FC_DL_GcdUdintCalc : UDINT
VAR_INPUT
    nA : UDINT := 0; // 左操作数 [脉冲 / 计数]，无符号 / the left operand, unsigned
    nB : UDINT := 0; // 右操作数 [脉冲 / 计数]，无符号 / the right operand, unsigned
END_VAR
VAR_OUTPUT
    nIter  : DINT;  // 迭代计数 [次]，供收敛审计 / the iteration count for the convergence audit
    bValid : BOOL;  // 结果可用 [-]（双零哨兵也是可用结果）/ the result usable, the zero sentinel is still usable
    eErr   : UDINT; // 错误码，0 = 正常 / the error code, zero is ok
    bError : BOOL;  // 故障标志（故障级码同拍置位，R45 配对）/ the fault flag raised with a fault level code
END_VAR
VAR
    nX   : UDINT := 0; // 迭代被除数工作副本 [脉冲 / 计数] / the dividend working copy of the iteration
    nY   : UDINT := 0; // 迭代除数工作副本 [脉冲 / 计数] / the divisor working copy of the iteration
    nRem : UDINT := 0; // 余数承接量 [脉冲 / 计数] / the remainder holder
END_VAR  // R64 结构补齐：VAR 段缺失的 END_VAR（门禁机械修复）
VAR CONSTANT
    DL_GCD_ZERO    : UDINT := 0;  // 无符号零常量 [脉冲 / 计数] / the unsigned zero constant
    DL_GCD_GUARDMAX: DINT   := 64; // WHILE 守卫计数上界 [次]（欧几里得迭代理论步数远小于此）/ the while guard ceiling, the euclid iteration converges far earlier
    DL_GCD_ZEROI   : DINT   := 0;  // 整型零常量 [次] / the integer zero constant
    DL_GCD_ONEI    : DINT   := 1;  // 整型一常量 [次] / the integer one constant
END_VAR

// 段 1｜返回值与全部出口预置安全值（R45 四段式第一段）/ segment 1, the preset of the return and all outlets
FC_DL_GcdUdintCalc := DL_GCD_ZERO; // 返回值预置 0 哨兵 / preset the return to the zero sentinel
nIter := DL_GCD_ZEROI; // 迭代计数预置零 [次] / preset the iteration count zero
bValid := FALSE; // 可用标志预置假 / preset the validity false
eErr := 16#0000_0000; // 错误码预置正常 / preset the code to ok
bError := FALSE; // 故障标志预置假 / preset the fault flag false
nX := DL_GCD_ZERO; // 被除数副本预置零 / preset the dividend copy zero
nY := DL_GCD_ZERO; // 除数副本预置零 / preset the divisor copy zero
nRem := DL_GCD_ZERO; // 余数承接量预置零 / preset the remainder holder zero

// 段 2｜双零哨兵（边界一：GCD(0,0) 无定义，信息级不置 bError）/ segment 2, the double zero sentinel
IF (nA = DL_GCD_ZERO) AND (nB = DL_GCD_ZERO) THEN // 双零入参 / both operands are zero
    eErr := 16#0001_0663; // 信息级：双零哨兵（R285）/ informational, the double zero sentinel
    bError := FALSE; // 信息级不置故障标志 / keep the fault flag false, this is informational
    bValid := TRUE; // 哨兵 0 是合法甄别结果 / the sentinel zero is a legit discernible result
    RETURN; // 早退，返回 0 / early return with zero
END_IF

// 段 3｜欧几里得迭代（边界二：MOD 除子 nY 由循环条件证明非零；边界三：守卫计数）/ segment 3, the euclid iteration with the proven divisor and the guard
nX := nA; // 被除数接管 [脉冲 / 计数] / take the dividend
nY := nB; // 除数接管 [脉冲 / 计数] / take the divisor
WHILE (nY <> DL_GCD_ZERO) AND (nIter < DL_GCD_GUARDMAX) DO // 除子非零且守卫未越限 / the divisor is nonzero and the guard is not exceeded
    nRem := nX MOD nY; // 余量（除子 nY 已由循环条件证明非零，除零不可达）/ the remainder, the divisor proven nonzero by the loop condition
    nX := nY; // 欧几里得步进：被除数取旧除数 / the euclid step, the dividend takes the old divisor
    nY := nRem; // 除数取余量 / the divisor takes the remainder
    nIter := nIter + DL_GCD_ONEI; // 迭代计数推进 [次] / advance the iteration count
END_WHILE

// 段 4｜守卫命中闸与统一出口（边界三）/ segment 4, the guard hit gate and the unified outlet
IF nY <> DL_GCD_ZERO THEN // 迭代因守卫越限退出（余量未收敛，平台异常路径）/ the loop exited by the guard with a nonzero remainder
    eErr := 16#0001_0664; // 故障级：守卫计数越限 / fault grade, the guard count exceeded
    bError := TRUE; // 同拍置故障标志（R45 配对）/ raise the fault flag on the same scan
    bValid := FALSE; // 结果不可用 / the result is not usable
    FC_DL_GcdUdintCalc := DL_GCD_ZERO; // 返回 0 哨兵（禁输出未收敛残值）/ return the zero sentinel, no unconverged residue
    RETURN; // 早退 / early return
END_IF
FC_DL_GcdUdintCalc := nX; // GCD 结果出口 [脉冲 / 计数]（nY 已收敛为 0，nX 即最大公约数）/ the gcd outlet with the converged value
bValid := TRUE; // 结果可用 / the result is usable
END_FUNCTION

(* ---- FC_DL_GearAddendumCircleCalc.st ---- *)
(*
  DL Factory R88 | FC_DL_GearAddendumCircleCalc
  功能：由模数/齿数/齿顶高系数算齿顶圆直径 da 与分度圆直径 d=m·z（da=d+2·ha*·m，标准齿 ha*=1）
  开源溯源：无（clean-room 自研，依据公开工艺公式 齿顶圆直径式 da=m·z+2·ha*·m，许可证=MIT，借鉴点=公式结构）
  规则：R1-R16 全遵守；R88 简单件标量形（纯标量入参出参，无循环体、无方法、无属性、无数组）
*)
FUNCTION FC_DL_GearAddendumCircleCalc : REAL
VAR_INPUT
    fModuleMm : REAL := 3.0; // 模数 m [mm] / module [mm]
    nTeeth : DINT := 20; // 齿数 z（整数入参，不可能为 NaN） [枚] / tooth count, integer input cannot be NaN [-]
    fAddFactor : REAL := 1.0; // 齿顶高系数 ha*（标准齿 1.0，短齿 0.8，长齿 1.2） [-] / addendum coefficient [-]
END_VAR
VAR_OUTPUT
    fDaMm : REAL; // 齿顶圆直径 da [mm] / addendum circle diameter [mm]
    fPitchDiaMm : REAL; // 分度圆直径 d [mm] / pitch circle diameter [mm]
END_VAR
VAR
    fTeeth : REAL; // 齿数实数化结果 [-] / tooth count converted to REAL [-]
    fAddendumMm : REAL; // 齿顶高 ha=ha*·m [mm] / addendum height [mm]
END_VAR

// 段 1｜出口预置
FC_DL_GearAddendumCircleCalc := -1.0; // 哨兵返回 -1（无效） [-] / sentinel return -1, invalid [-]
fDaMm := 0.0; // 齿顶圆直径预置零 [mm] / addendum diameter preset zero [mm]
fPitchDiaMm := 0.0; // 分度圆直径预置零 [mm] / pitch diameter preset zero [mm]
fTeeth := 0.0; // 齿数实数预置零 [-] / real teeth preset zero [-]
fAddendumMm := 0.0; // 齿顶高预置零 [mm] / addendum preset zero [mm]

// 段 2｜非有限拦截 + 域闸
IF NOT (fModuleMm > -1.0E30 AND fModuleMm < 1.0E30) OR NOT (fAddFactor > -1.0E30 AND fAddFactor < 1.0E30) THEN
    RETURN; // 模数/齿顶高系数任一非有限即拒算 [-] / any non finite input rejected [-]
END_IF
IF fModuleMm < 1.0E-9 THEN
    RETURN; // 模数正域闸 [mm] / positive module gate [mm]
END_IF
IF fAddFactor < 0.4 OR fAddFactor > 1.6 THEN
    RETURN; // 齿顶高系数工程域闸（远离 0 防退化齿形） [-] / addendum coefficient domain gate [-]
END_IF
IF nTeeth < 1 THEN
    RETURN; // 齿数下限闸（整数域，无 NaN 可能，仅做范围拦截） [枚] / tooth count lower gate [-]
END_IF

// 段 3｜计算
fTeeth := DINT_TO_REAL(nTeeth); // DINT→REAL 标准转换函数（R10 禁构造函数式） [-] / standard conversion function (R10) [-]
fAddendumMm := fAddFactor * fModuleMm; // 无量纲 × mm = mm，ha=ha*·m / [-] × [mm] = [mm]
fPitchDiaMm := fModuleMm * fTeeth; // mm × 无量纲 = mm，d=m·z / [mm] × [-] = [mm]
fDaMm := fPitchDiaMm + 2.0 * fAddendumMm; // mm + mm = mm，da=d+2·ha=m·z+2·ha*·m [mm] / [mm]

// 段 4｜判定与饱和
IF fDaMm <= fPitchDiaMm THEN
    RETURN; // 结构自洽闸：齿顶圆必须严格大于分度圆 [mm] / structural check da > d [mm]
END_IF

// 段 5｜出口自检
IF NOT (fDaMm > -1.0E30 AND fDaMm < 1.0E30) OR fDaMm < 1.0E-9 THEN
    RETURN; // 出口自检：齿顶圆有限且为正，否则退回哨兵 [mm] / exit self-check on da [mm]
END_IF
FC_DL_GearAddendumCircleCalc := fDaMm; // 返回齿顶圆直径 [mm] / return the addendum diameter [mm]
END_FUNCTION

(* ---- FC_DL_GearBaseCircleCalc.st ---- *)
(*
  DL Factory R88 | FC_DL_GearBaseCircleCalc
  功能：由模数/齿数/压力角算基圆直径 db=m·z·cosα，压力角由角度制按 π/180 换算弧度
  开源溯源：无（clean-room 自研，依据公开工艺公式 基圆直径式 db=m·z·cosα，许可证=MIT，借鉴点=公式结构）
  规则：R1-R16 全遵守；R88 简单件标量形（纯标量入参出参，无循环体、无方法、无属性、无数组）
*)
FUNCTION FC_DL_GearBaseCircleCalc : REAL
VAR_INPUT
    fModuleMm : REAL := 3.0; // 模数 m [mm] / module [mm]
    nTeeth : DINT := 20; // 齿数 z（整数入参，无 NaN 可能） [枚] / tooth count, integer input [-]
    fPressureDeg : REAL := 20.0; // 分度圆压力角 α（度制，域闸 10~30） [°] / pressure angle in degrees [-]
END_VAR
VAR_OUTPUT
    fDbMm : REAL; // 基圆直径 db [mm] / base circle diameter [mm]
    fPitchDiaMm : REAL; // 分度圆直径 d=m·z [mm] / pitch circle diameter [mm]
END_VAR
VAR
    fTeeth : REAL; // 齿数实数化结果 [-] / tooth count converted to REAL [-]
    fAlphaRad : REAL; // 压力角弧度值 [rad] / pressure angle in radians [rad]
    fCosAlpha : REAL; // 压力角余弦（缓存，避免重算） [-] / cosine of the pressure angle [-]
END_VAR

// 段 1｜出口预置
FC_DL_GearBaseCircleCalc := -1.0; // 哨兵返回 -1（无效） [-] / sentinel return -1, invalid [-]
fDbMm := 0.0; // 基圆直径预置零 [mm] / base diameter preset zero [mm]
fPitchDiaMm := 0.0; // 分度圆直径预置零 [mm] / pitch diameter preset zero [mm]
fTeeth := 0.0; // 齿数实数预置零 [-] / real teeth preset zero [-]
fAlphaRad := 0.0; // 弧度预置零 [rad] / radians preset zero [rad]
fCosAlpha := 0.0; // 余弦预置零 [-] / cosine preset zero [-]

// 段 2｜非有限拦截 + 域闸
IF NOT (fModuleMm > -1.0E30 AND fModuleMm < 1.0E30) OR NOT (fPressureDeg > -1.0E30 AND fPressureDeg < 1.0E30) THEN
    RETURN; // 模数/压力角任一非有限即拒算 [-] / any non finite input rejected [-]
END_IF
IF fModuleMm < 1.0E-9 THEN
    RETURN; // 模数正域闸 [mm] / positive module gate [mm]
END_IF
IF fPressureDeg <= 10.0 OR fPressureDeg >= 30.0 THEN
    RETURN; // 压力角开区间域闸 (10°,30°)：趋零则基圆退化为分度圆 [°] / open interval gate on alpha [deg]
END_IF
IF nTeeth < 1 THEN
    RETURN; // 齿数下限闸（整数域，仅做范围拦截） [枚] / tooth count lower gate [-]
END_IF

// 段 3｜计算
fTeeth := DINT_TO_REAL(nTeeth); // DINT→REAL 标准转换函数（R10） [-] / standard conversion function (R10) [-]
fAlphaRad := fPressureDeg * 0.0174532925; // 度 × (π/180) = rad，换算常数 0.0174532925 [rad] / degrees to radians [rad]
fCosAlpha := COS(fAlphaRad); // 无量纲 [-] / dimensionless cosine [-]
fPitchDiaMm := fModuleMm * fTeeth; // mm × 无量纲 = mm，d=m·z / [mm] × [-] = [mm]
fDbMm := fPitchDiaMm * fCosAlpha; // mm × 无量纲 = mm，db=d·cosα / [mm] × [-] = [mm]

// 段 4｜判定与饱和
IF fDbMm <= 0.0 THEN
    RETURN; // 结果闸：基圆直径必须为正（cosα 在 (10°,30°) 内恒正） [mm] / base diameter must be positive [mm]
END_IF
IF fDbMm >= fPitchDiaMm THEN
    RETURN; // 结构自洽闸：基圆必须小于分度圆（cosα<1） [mm] / structural check db < d [mm]
END_IF

// 段 5｜出口自检
IF NOT (fDbMm > -1.0E30 AND fDbMm < 1.0E30) THEN
    RETURN; // 出口自检：结果非有限即退回哨兵 [mm] / exit self-check on finiteness [mm]
END_IF
FC_DL_GearBaseCircleCalc := fDbMm; // 返回基圆直径 [mm] / return the base circle diameter [mm]
END_FUNCTION
